(* IEC 61131-3 sources: daoli-st-library/DL_Algo (part 23) *)

(* ---- FB_DL_TriangleGenerator.st ---- *)
(*
  FB_DL_TriangleGenerator  —  三角波发生（相位连续 + 幅值/频率引脚化）/ Triangle wave generator
  分类 Category : DL_Algo
  码位 Code     : 16#02_3_87
  段位说明      : 86 格由 FB_DL_FrequencyGenerator 启用，本件启用相邻 87 格（一件一码）
  版本 Version  : 1.0.0
  来源 Source   : t2-1-lgf-siggen — 信号发生族第三基本波形（Sine/Sawtooth 同族）
  溯源 Origin   : clean-room 实现，相位累加三角波为公开经典方法，未复制任何源码行
  功能 Function : 1) 三角波发生：相位累加器在 [0,1) 内推进，方向标志交替升/降，
                  归一化输出 fNorm ∈ [0,1]，工程输出 fOut = fOffset + fAmplitude * (2*fNorm − 1)；
                  2) bPhaseReset 上升沿强制相位归零且方向置升（多路同相启动）；
                  3) fFreqHz = 0 时冻结在当前相位值（静止保持，不清输出）；
                  4) 波形形状按矩阵组纪律独立成件，明文禁用 eWaveform 枚举合并
                  （与 FB_DL_SineGenerator / 锯齿族分工，本件只做三角）。
  边界 Boundary : ① 幅值允许负值（输出相位反转语义：负幅值 = 倒相），非有限防御保持上次有效值；
                  ② 偏移 fOffset 非有限防御保持上次有效值；首扫按默认值；
                  ③ 无 TON/边沿实例：相位累加器法，任务周期由调用方经 tSampleTime 注入，
                  < T#10MS 钳位（与 FB_DL_RateLimiter 同口径）；
                  ④ 频率上限钳位（奈奎斯特防御）：高于任务频率一半时波形失真，越限按上限执行并置信息码；
                  ⑤ 方向切换在同一拍完成：fPhase >= 1 时先翻转方向再截去进位，避免相位突变尖峰。
  依赖 Depends  : 仅 Standard.library；与 FB_DL_SineGenerator（已注册）仅引脚口径对齐，不实例化
  码表 Error codes（本件格 02_3_87，子码步进 +0x100）:
    16#0002_0187 信息级：频率越上限已钳位（奈奎斯特防御，输出按钳后频率执行）
    16#0002_0287 信息级：相位复位沿生效（fPhase 归零、方向置升）
    16#0002_0387 信息级：非有限参数防御触发（保持上次有效值继续运行）

  修订历史 Revision :
    2026-11-19  v1.0.0  R39 首版（批次 1 · 序号 5）
*)

FUNCTION_BLOCK FB_DL_TriangleGenerator
VAR_INPUT
    bEnable     : BOOL := FALSE;      // 使能，FALSE 时冻结相位与输出 [-] / Enable, FALSE freezes phase and output
    fFreqHz     : REAL := 1.0;        // 目标频率 [Hz]，域 (0, 上限]，越限钳位 / Target frequency [Hz], clamped
    fAmplitude  : REAL := 100.0;      // 幅值 [EU]，可负（倒相语义），非有限保持 / Amplitude [EU], negative inverts phase
    fOffset     : REAL := 0.0;        // 直流偏移 [EU]，非有限保持 / DC offset [EU]
    bPhaseReset : BOOL := FALSE;      // 相位复位，上升沿相位归零、方向置升 / Phase reset, rising edge zeroes phase
    tSampleTime : TIME := T#100MS;    // 任务周期注入 [ms]，< T#10MS 钳位 / Task cycle time injected by caller
END_VAR
VAR_OUTPUT
    fOut        : REAL;               // 三角波工程输出 [EU] / Triangle engineering output [EU]
    fNormOut    : REAL;               // 归一化输出 [无量纲 0..1]，0 = 谷 / Normalized output, 0 = valley
    bRising     : BOOL;               // 本拍处于上升半周 [-] / Currently in the rising half-cycle
    uCycleCnt   : UDINT;              // 完整周期计数 [次]，降→升切换计一次，饱和 / Full cycle count, saturating
    bError      : BOOL;               // 故障标志，本件全信息级恒 FALSE（R21：信息级码不置故障）[-] / Fault flag, always FALSE, all codes info level
    uErrorId    : UDINT;              // 事件码，0 = 无事件（本件码均瞬时逐拍重算）/ Event code, transient, recomputed each scan
END_VAR
VAR
    rtPhaseReset : R_TRIG;            // 相位复位沿实例，主体首部无条件刷新 / Phase reset edge instance
    _fPhase      : REAL := 0.0;       // 内部相位累加器 [无量纲 0..1) / Internal phase accumulator
    _bUp         : BOOL := TRUE;      // 内部方向标志，TRUE = 升半周 / Internal direction flag, TRUE = rising
    _fFreqEff    : REAL := 1.0;       // 钳位后的生效频率 [Hz] / Clamped effective frequency
    _fAmpEff     : REAL := 100.0;     // 生效幅值 [EU] / Effective amplitude
    _fOffEff     : REAL := 0.0;       // 生效偏移 [EU] / Effective offset
    _fDt         : REAL := 0.1;       // 生效任务周期 [s] / Effective cycle time in seconds
    _fFreqLast   : REAL := 1.0;       // 上次有效频率保持载体 [Hz] / Last valid frequency hold carrier
    _fAmpLast    : REAL := 100.0;     // 上次有效幅值保持载体 [EU] / Last valid amplitude hold carrier
    _fOffLast    : REAL := 0.0;       // 上次有效偏移保持载体 [EU] / Last valid offset hold carrier
    _fNorm       : REAL := 0.0;       // 归一化中间量 [无量纲 0..1] / Normalized working value
    _bDefend     : BOOL;              // 本拍非有限防御触发标志 / Non-finite defense triggered this cycle
END_VAR
VAR CONSTANT
    DL_TG_DT_MIN     : TIME := T#10MS;      // 任务周期下限钳位 [ms] / Cycle time lower clamp
    DL_TG_FREQ_MAX   : REAL := 5.0;         // 频率组态上限（奈奎斯特防御，按 100ms 任务口径）[Hz] / Frequency configuration bound
    DL_TG_INF_CAP    : REAL := 1.0E30;      // 非有限值筛查幅值上限 / Non-finite magnitude screening cap
    DL_TG_CNT_MAX    : UDINT := 16#FFFF_FFFE;  // 周期计数饱和上限 [次] / Cycle count saturation bound
END_VAR

(* —— 段 0：边沿实例无条件周期刷新（R7 红线：严禁置于 IF/CASE 分支内） —— *)
rtPhaseReset(CLK := bPhaseReset);       // 相位复位沿刷新，每拍必调

(* —— 段 1：单拍量预清零 —— *)
uErrorId := 16#0000_0000;               // 事件码每拍重算（本件全信息级）
_bDefend := FALSE;                      // 防御标志预清零

(* —— 段 2：非有限防御与参数钳位（NaN/Inf 保持上次有效值） —— *)
IF (fFreqHz <> fFreqHz) OR (ABS(fFreqHz) > DL_TG_INF_CAP) OR ((fFreqHz - fFreqHz) <> 0.0) THEN
    _fFreqEff := _fFreqLast;            // 频率非有限：保持上次有效
    _bDefend := TRUE;
ELSE
    _fFreqLast := fFreqHz;
    IF fFreqHz < 0.0 THEN
        _fFreqEff := 0.0;               // 负频率钳零（冻结在当前相位值）
    ELSIF fFreqHz > DL_TG_FREQ_MAX THEN
        _fFreqEff := DL_TG_FREQ_MAX;    // 越上限钳位（奈奎斯特防御）
        uErrorId := 16#0002_0187;       // 信息级：频率已钳位
    ELSE
        _fFreqEff := fFreqHz;           // 域内直通
    END_IF
END_IF
IF (fAmplitude <> fAmplitude) OR (ABS(fAmplitude) > DL_TG_INF_CAP) OR ((fAmplitude - fAmplitude) <> 0.0) THEN
    _fAmpEff := _fAmpLast;              // 幅值非有限：保持上次有效
    _bDefend := TRUE;
ELSE
    _fAmpLast := fAmplitude;
    _fAmpEff := fAmplitude;             // 幅值允许负值（倒相语义），不钳位
END_IF
IF (fOffset <> fOffset) OR (ABS(fOffset) > DL_TG_INF_CAP) OR ((fOffset - fOffset) <> 0.0) THEN
    _fOffEff := _fOffLast;              // 偏移非有限：保持上次有效
    _bDefend := TRUE;
ELSE
    _fOffLast := fOffset;
    _fOffEff := fOffset;                // 偏移直通
END_IF
IF _bDefend THEN
    uErrorId := 16#0002_0387;           // 信息级：非有限防御触发（覆盖钳位码，防御码优先）
END_IF

(* —— 段 3：任务周期换算（与 FB_DL_RateLimiter 同口径：< T#10MS 钳位） —— *)
IF tSampleTime < DL_TG_DT_MIN THEN
    _fDt := 0.01;                       // 非法周期钳位 0.01 s
ELSE
    _fDt := TIME_TO_REAL(tSampleTime) / 1000.0;   // TIME 换算秒（显式标准转换）
END_IF

(* —— 段 4：相位复位沿（先于推进处理） —— *)
IF rtPhaseReset.Q THEN
    _fPhase := 0.0;                     // 相位归零
    _bUp := TRUE;                       // 方向置升
    uErrorId := 16#0002_0287;           // 信息级：相位复位生效（覆盖防御码，复位意图优先显式）
END_IF

(* —— 段 5：相位推进与方向翻转（失能冻结；频率 0 冻结在当前值） —— *)
IF bEnable AND (_fFreqEff > 0.0) THEN
    _fPhase := _fPhase + _fFreqEff * _fDt;      // 相位推进 = 频率 × 周期
    IF _fPhase >= 1.0 THEN
        _fPhase := _fPhase - 1.0;               // 截去进位（同拍完成，避免相位突变尖峰）
        IF _bUp THEN
            _bUp := FALSE;                      // 升满翻降（峰点换向）
        ELSE
            _bUp := TRUE;                       // 降满翻升（谷点换向）
            uCycleCnt := uCycleCnt + 1;         // 完整周期计数（降→升切换口径）
            IF uCycleCnt >= DL_TG_CNT_MAX THEN
                uCycleCnt := DL_TG_CNT_MAX;     // 计数饱和防回绕
            END_IF
        END_IF
        IF _fPhase >= 1.0 THEN
            _fPhase := 0.0;                     // 极端钳位兜底（频率越限多周回绕）
        END_IF
    END_IF
END_IF

(* —— 段 6：波形合成（升半周 fNorm = fPhase，降半周 fNorm = 1 − fPhase） —— *)
IF _bUp THEN
    _fNorm := _fPhase;                          // 上升半周：归一化随相位升
ELSE
    _fNorm := 1.0 - _fPhase;                    // 下降半周：归一化随相位降
END_IF
fNormOut := _fNorm;                             // 归一化镜像输出
fOut := _fOffEff + _fAmpEff * (2.0 * _fNorm - 1.0);   // 工程输出 = 偏移 + 幅值 ×（2·归一化 − 1）
bRising := _bUp AND bEnable;                    // 上升半周指示（失能时恒 FALSE）
bError := FALSE;                                // 本件全信息级：故障位恒 FALSE（R21）

END_FUNCTION_BLOCK

(* ---- FB_DL_TwoDofPid.st ---- *)
(*
  ==================================================================
  组件名 Component  : FB_DL_TwoDofPid
  分类   Category   : DL_Algo
  复杂度 Complexity  : cx4
  版本   Version    : 1.0.1
  功能   Purpose    : 二自由度 PID（设定值加权 beta / gamma），位置式：
                      u = Kp·(beta·sp - pv) + I + Kp·Td·(gamma·dsp/dt - dpv/dt)（滤后）。
                      积分作用于全误差 (sp - pv)；微分先行经 nFilter 一阶低通；
                      抗积分饱和（输出限幅方向与误差同向时停积分）；手动/自动
                      无扰切换（手动相把积分项跟踪为 fManOut - P - D）。
  来源   Source     : t2-5-modpid（参数域 beta / gamma）
  溯源   Origin     : IEC 61131-3 标准语义的道莅防御性实现；二自由度 PID 结构为
                      公开控制理论结果（Araki 参考跟踪 / 扰动抑制双自由度组织），
                      clean-room 自研实现，未复制任何闭源代码行。
  平台   Platform   : 纯 IEC 61131-3（LREAL 运算，无私有库、无幂运算符）
  作者   Author     : 道莅代码库 · PLC 编程专家（R56）
  ------------------------------------------------------------------
  边界 Boundary     :
                      一 本件只算控制器输出，不驱动执行器、不做自整定（属主边界）；
                      二 同拍双窗说明（R100）：本件无同拍双 TON 结构，微分滤波为一阶
                         差分实现，无定时器实例；
                      三 fTi <= 0 时积分项关闭（纯 PD 口径），fTd <= 0 时微分项关闭；
                      四 bInvalid = TRUE 时输出冻结保持末值（R191 显式声明，降级不静默）；
                      五 故障锁存（组态非法）解除路径 = bReset 上升沿（唯一路径，R188）；
                      六 无全局变量、无外部变量声明、无物理地址寻址、无定时器实例。
  输出契约 Output contract:
                      fOut 恒被钳在 [fOutMin, fOutMax]；bSatHi / bSatLo 为本拍限幅指示；
                      eFault 为锁存回放（eCfgIllegal 组态非法 / eInputBad 本拍输入非有限）。
  修订记录 Revision  :
    2026-11-20  v1.0.0  R56 首版（批 2 · 序号 8）
    2026-11-21  v1.0.1  R57 返修：手动相入口补 fManOut 有限性闸，无效拍冻结早退不进跟踪式
  ==================================================================
*)

TYPE E_DL_TdpFault :
(
    eNone     := 0, // 无成因 / no cause
    eCfgIllegal := 1, // 组态非法：增益或限幅越域（故障级，与 bError 配对）/ illegal config, gain or limit out of domain
    eInputBad := 2  // 本拍设定值或过程量非有限（信息级，输出冻结保持）/ the setpoint or process value is non finite this scan, the output holds frozen
);
END_TYPE

FUNCTION_BLOCK FB_DL_TwoDofPid
VAR_INPUT
    bAuto    : BOOL := TRUE;     // 自动模式，假 = 手动（无扰切换）[-] / auto mode, false is manual with a bumpless transfer
    bReset   : BOOL := FALSE;    // 复位上升沿清故障锁存与积分 [-] / reset rising edge clears the fault latch and the integral
    fSp      : LREAL := 0.0;     // 设定值 [工程单位] / setpoint [engineering unit]
    fPv      : LREAL := 0.0;     // 过程量实测 [工程单位] / measured process value [engineering unit]
    fManOut  : LREAL := 0.0;     // 手动输出值 [工程单位] / manual output value [engineering unit]
    fKp      : LREAL := 1.0;     // 比例增益，域 大于零 / proportional gain, domain above zero
    fTi      : LREAL := 10.0;    // 积分时间 [秒]，0 = 积分关闭 / integral time [second], zero disables the integral
    fTd      : LREAL := 0.0;     // 微分时间 [秒]，0 = 微分关闭 / derivative time [second], zero disables the derivative
    fBeta    : LREAL := 1.0;     // 设定值比例加权（抑超调自由度），域 0..1 / setpoint proportional weight [dimensionless], domain zero to one
    fGamma   : LREAL := 0.0;     // 设定值微分加权，域 0..1 / setpoint derivative weight, domain zero to one
    nFilter  : INT := 10;        // 微分低通系数 n（Td/n 为滤波时间），域 1..100 / derivative low pass coefficient n, domain one to one hundred
    fOutMin  : LREAL := 0.0;     // 输出下限 [工程单位] / output floor [engineering unit]
    fOutMax  : LREAL := 100.0;   // 输出上限 [工程单位]，域 大于下限 / output ceiling [engineering unit], above the floor
    fDtS     : LREAL := 0.01;    // 调用周期 [秒]，域 大于零 / call period [second], domain above zero
END_VAR
VAR_OUTPUT
    fOut     : LREAL := 0.0;   // 控制器输出 [工程单位] / controller output [engineering unit]
    bSatHi   : BOOL := FALSE;  // 本拍输出顶上限 [-] / the output hit the ceiling this scan
    bSatLo   : BOOL := FALSE;  // 本拍触下限 [-] / the output hit the floor this scan
    bInvalid : BOOL := FALSE;  // 本拍输出无效（冻结保持末值）[-] / the outlet is void this scan, the last value holds frozen
    eFault   : E_DL_TdpFault := E_DL_TdpFault.eNone; // 成因出口，锁存回放 [枚举] / cause outlet replayed from the latch [enum]
    bError   : BOOL := FALSE;  // 故障锁存标志 [-] / fault latch flag
END_VAR
VAR
    rtReset  : R_TRIG;  // 复位沿检测，段 0 无条件刷新 / reset edge, refreshed unconditionally in segment zero
    _eFaulC  : E_DL_TdpFault := E_DL_TdpFault.eNone; // 故障级成因，锁存至复位沿 / fault cause, latched until the reset edge
    _bFault  : BOOL := FALSE; // 故障锁存位 [-] / fault latch bit
    _bInit   : BOOL := FALSE; // 首扫初始化完成标志（R310）/ first scan initialisation flag
    _bInOk   : BOOL := FALSE; // 本拍 sp / pv 均有限 [-] / both sp and pv are finite this scan
    _fI      : LREAL := 0.0;  // 积分项保持量 [工程单位] / the integral term holder [engineering unit]
    _fDfilt  : LREAL := 0.0;  // 微分滤波保持量 [工程单位] / the derivative filter holder [engineering unit]
    _fPvPrev : LREAL := 0.0;  // 上拍过程量快照 [工程单位] / previous scan process value snapshot [engineering unit]
    _fSpPrev : LREAL := 0.0;  // 上拍设定值快照 [工程单位] / previous scan setpoint snapshot [engineering unit]
    _fP      : LREAL := 0.0;  // 本拍比例项 [工程单位] / the proportional term this scan [engineering unit]
    _fDraw   : LREAL := 0.0;  // 微分原始量 [工程单位] / the raw derivative term [engineering unit]
    _fE      : LREAL := 0.0;  // 全误差（sp - pv）[工程单位] / the full error [engineering unit]
    _fUPre   : LREAL := 0.0;  // 限幅前输出 [工程单位] / the pre clamp output [engineering unit]
    _fFiltB  : LREAL := 0.0;  // 微分滤波权（dt/(dt+Td/n)）[无量纲] / the derivative filter weight
END_VAR

// 段 0｜沿检测无条件周期刷新（禁入分支）/ segment 0, unconditional refresh of the edge detector
rtReset(CLK := bReset); // 复位沿无条件刷新 / unconditional refresh of the reset edge

// 段 1｜首扫初始化（R310）：快照与积分从确定起点起步 / segment 1, first scan initialisation
IF NOT _bInit THEN // 首扫一拍 / the very first scan
    _bInit := TRUE; // 置首扫完成标志 / raise the first scan flag
    _eFaulC := E_DL_TdpFault.eNone; // 故障级成因清零 / clear the fault cause
    _bFault := FALSE; // 故障锁存清零 / clear the fault latch
    _fI := 0.0; // 积分项清零 / clear the integral term
    _fDfilt := 0.0; // 微分滤波清零 / clear the derivative filter
    _fPvPrev := fPv; // 快照取当拍 / the snapshot takes this scan
    _fSpPrev := fSp; // 快照取当拍 / the snapshot takes this scan
END_IF

// 段 2｜复位沿作用域：清锁存 / 清积分与滤波（快照同步归位，三项逐项声明）/ segment 2, reset edge scope declared item by item
IF rtReset.Q THEN // 复位沿 / the reset edge
    _bFault := FALSE; // 作用域一：清故障锁存 / scope one, clear the fault latch
    _eFaulC := E_DL_TdpFault.eNone; // 作用域一：清故障级成因 / scope one, clear the fault cause
    _fI := 0.0; // 作用域二：清积分项 / scope two, clear the integral term
    _fDfilt := 0.0; // 作用域二：清微分滤波 / scope two, clear the derivative filter
    _fPvPrev := fPv; // 作用域三：快照归位 / scope three, the snapshot parks
    _fSpPrev := fSp; // 作用域三：快照归位 / scope three, the snapshot parks
END_IF

// 段 3｜组态域闸（R151 全覆盖）/ segment 3, configuration domain gate over every parameter pin
IF (fKp <= 0.0) OR (fKp <> fKp) OR ((fKp - fKp) <> (fKp - fKp)) OR (fTi < 0.0) OR (fTi <> fTi) OR (fTd < 0.0) OR (fTd <> fTd) OR (fBeta < 0.0) OR (fBeta > 1.0) OR (fBeta <> fBeta) OR (fGamma < 0.0) OR (fGamma > 1.0) OR (fGamma <> fGamma) OR (nFilter < 1) OR (nFilter > 100) OR (fOutMax <= fOutMin) OR (fOutMax <> fOutMax) OR (fDtS <= 0.0) OR (fDtS <> fDtS) THEN // 任一参数越域或非有限 / any parameter out of domain or non finite
    IF (NOT _bFault) AND (_eFaulC = E_DL_TdpFault.eNone) THEN // 未锁存才迁移（防同拍抹除）/ migrate only while unlatched
        _bFault := TRUE; // 置故障锁存 / raise the fault latch
        _eFaulC := E_DL_TdpFault.eCfgIllegal; // 故障级成因（R45 配对 bError）/ the fault cause paired with bError
    END_IF
END_IF

// 段 4｜输入有限性闸与冻结语义 / segment 4, the input finiteness gate and the frozen semantics
_bInOk := (fSp = fSp) AND ((fSp - fSp) = (fSp - fSp)) AND (fPv = fPv) AND ((fPv - fPv) = (fPv - fPv)); // sp / pv 有限性 / finiteness of sp and pv

// 段 5｜无扰切换：手动相把积分项跟踪为 fManOut - P - D / segment 5, the bumpless transfer, the manual phase tracks the integral
IF NOT bAuto THEN // 手动相 / the manual phase
    IF (fManOut <> fManOut) OR ((fManOut - fManOut) <> (fManOut - fManOut)) THEN // 手动输出非有限（x<>x 判 NaN，x-x<>x-x 判 Inf，v1.0.1 返修）/ the manual output is non finite (v1.0.1 fix)
        IF NOT _bFault THEN // 故障锁存优先回放，信息级不覆盖故障码 / the fault latch replays first, an informational cause never overwrites a fault code
            _eFaulC := E_DL_TdpFault.eInputBad; // 信息级成因（R45 不配对 bError）/ the informational cause, not paired with bError
        END_IF
        bInvalid := TRUE; // 置无效标志 / raise the invalid flag
        bSatHi := FALSE; // 限幅指示为假 / the saturation flags are false
        bSatLo := FALSE; // 限幅指示为假 / the saturation flags are false
        eFault := _eFaulC; // 成因出口锁存回放 / the cause outlet replayed from the latch
        bError := _bFault; // 故障标志与锁存位同源 / the fault flag shares the latch source
        _fPvPrev := fPv; // 快照推进（防恢复时微分踢）/ advance the snapshot against a derivative kick
        _fSpPrev := fSp; // 快照推进 / advance the snapshot
        RETURN; // 早退，fOut 冻结保持末值，不进跟踪式（R191 已声明）/ early return, fOut holds frozen, no tracking (R191 declared)
    END_IF
    _fP := fKp * (fBeta * fSp - fPv); // 比例项同口径计算（为跟踪做准备）/ the proportional term for the tracking base
    _fI := fManOut - _fP - _fDfilt; // 积分项跟踪，自动恢复时无扰 / the integral tracks for a bumpless auto resume
    fOut := fManOut; // 手动输出直通 / the manual output passes through
    IF fOut > fOutMax THEN // 手动输出上钳 / clamp the manual output high
        fOut := fOutMax; // 钳到上限 / clamp to the ceiling
    ELSIF fOut < fOutMin THEN // 手动输出下钳 / clamp the manual output low
        fOut := fOutMin; // 钳到下限 / clamp to the floor
    END_IF
    bSatHi := FALSE; // 手动相限幅指示为假 / the saturation flags are false in manual
    bSatLo := FALSE; // 手动相限幅指示为假 / the saturation flags are false in manual
    bInvalid := (NOT _bInOk) OR _bFault; // 有效性随输入与锁存 / the validity follows the input and the latch
    eFault := _eFaulC; // 成因出口锁存回放 / the cause outlet replayed from the latch
    bError := _bFault; // 故障标志与锁存位同源 / the fault flag shares the latch source
    _fPvPrev := fPv; // 快照推进 / advance the snapshot
    _fSpPrev := fSp; // 快照推进 / advance the snapshot
    RETURN; // 手动相早退（出口段已完整施加，R94）/ the manual phase early return with a complete outlet
END_IF

// 段 6｜自动相：无效输入冻结保持 / segment 6, the auto phase, a void input holds frozen
IF (NOT _bInOk) OR _bFault THEN // 输入无效或故障锁存 / the input is void or faulted
    IF (NOT _bInOk) AND (NOT _bFault) THEN // 输入缺陷才记信息级成因（不覆盖故障码）/ only an input defect records the informational cause, never over a fault latch
        _eFaulC := E_DL_TdpFault.eInputBad; // 信息级成因，每拍重算 / the informational cause, recomputed every scan
    END_IF
    bInvalid := TRUE; // 置无效标志 / raise the invalid flag
    bSatHi := FALSE; // 限幅指示为假 / the saturation flags are false
    bSatLo := FALSE; // 限幅指示为假 / the saturation flags are false
    eFault := _eFaulC; // 成因出口锁存回放 / the cause outlet replayed from the latch
    bError := _bFault; // 故障标志与锁存位同源 / the fault flag shares the latch source
    _fPvPrev := fPv; // 快照推进（防恢复时微分踢）/ advance the snapshot against a derivative kick
    _fSpPrev := fSp; // 快照推进 / advance the snapshot
    RETURN; // 早退，fOut 冻结保持末值（R191 已在头注释声明）/ early return, fOut holds frozen per the declared semantics
END_IF

// 段 7｜比例与微分先行（幂次无，显式乘法）/ segment 7, the proportional and the derivative lead terms
_fE := fSp - fPv; // 全误差 / the full error
_fP := fKp * (fBeta * fSp - fPv); // 加权比例项 / the weighted proportional term
IF fTd > 0.0 THEN // 微分开启 / the derivative is on
    _fDraw := fTd * (fGamma * (fSp - _fSpPrev) - (fPv - _fPvPrev)) / fDtS; // 加权微分原始量，除子为周期已证大于零 / the weighted raw derivative, the divisor is the proven period
    _fFiltB := fDtS / (fDtS + fTd / INT_TO_LREAL(nFilter)); // 一阶低通权，除子已证大于零 / the first order weight with a proven divisor
    _fDfilt := _fDfilt + _fFiltB * (_fDraw - _fDfilt); // 微分低通推进 / advance the derivative low pass
ELSE // 微分关闭 / the derivative is off
    _fDfilt := 0.0; // 微分项归零 / the derivative term is zeroed
END_IF

// 段 8｜积分与抗饱和：先算限幅前输出，再按方向条件积分 / segment 8, the integral with anti windup, the clamp direction gates the accumulation
_fUPre := _fP + _fI + _fDfilt; // 限幅前输出 / the pre clamp output
IF (fTi > 0.0) THEN // 积分开启 / the integral is on
    IF NOT ((_fUPre > fOutMax) AND (_fE > 0.0)) AND NOT ((_fUPre < fOutMin) AND (_fE < 0.0)) THEN // 输出未沿误差方向饱和才积分（抗 windup）/ the integration only runs when the output is not saturated in the error direction
        _fI := _fI + (fKp / fTi) * _fE * fDtS; // 积分推进，除子为积分时间已证大于零 / the integral step with the proven divisor
    END_IF
END_IF
_fUPre := _fP + _fI + _fDfilt; // 积分后重算限幅前输出 / recompute after the integral

// 段 9｜限幅与限幅指示 / segment 9, the clamp and the saturation flags
bSatHi := FALSE; // 限幅指示预置假 / preset the saturation flags to false
bSatLo := FALSE; // 限幅指示预置假 / preset the saturation flags to false
IF _fUPre > fOutMax THEN // 顶上限 / above the ceiling
    fOut := fOutMax; // 钳到上限 / clamp to the ceiling
    bSatHi := TRUE; // 置顶上限指示 / raise the ceiling flag
ELSIF _fUPre < fOutMin THEN // 触下限 / below the floor
    fOut := fOutMin; // 钳到下限 / clamp to the floor
    bSatLo := TRUE; // 置触下限指示 / raise the floor flag
ELSE // 域内 / inside the domain
    fOut := _fUPre; // 直接出口 / straight to the outlet
END_IF

// 段 10｜快照推进与统一出口 / segment 10, the snapshot advance and the unified outlet
_fPvPrev := fPv; // 过程量快照推进 / advance the process snapshot
_fSpPrev := fSp; // 设定值快照推进 / advance the setpoint snapshot
IF (_eFaulC = E_DL_TdpFault.eInputBad) AND (NOT _bFault) THEN // 输入已恢复 / the input has recovered
    _eFaulC := E_DL_TdpFault.eNone; // 信息级成因随恢复撤销 / the informational cause is revoked on recovery
END_IF
bInvalid := FALSE; // 自动有效拍 / the valid auto scan
eFault := _eFaulC; // 成因出口锁存回放 / the cause outlet replayed from the latch
bError := _bFault; // 故障标志与锁存位同源 / the fault flag shares the latch source
END_FUNCTION_BLOCK

(* ---- FB_DL_UvDoseCtrl.st ---- *)
(*
  ==================================================================
  组件名 Component  : FB_DL_UvDoseCtrl
  分类   Category   : DL_Algo
  复杂度 Complexity  : cx5
  版本   Version    : 1.0.0
  功能   Purpose    : UV 剂量控制。剂量 = 光强 × 曝晒时间（D = ∫I·kLamp·dt），
                      按剩余剂量误差 PI 闭环调光强输出（0..100%），累计达目标置
                      bDoseDone 单拍脉冲；灯管老化补偿系数 kLamp 外部给定；光强
                      非有限 / 负值闸；累计溢出保护；满输出长期照度不足判
                      eLampWeak；过冲超容差判 eDoseOvershoot。
  来源   Source     : 自研线（公开物理定义：剂量 = 强度 × 时间积分）
  溯源   Origin     : IEC 61131-3 标准语义的道莅防御性实现；UV 剂量定义为公开
                      光化学语义，clean-room 自研实现，未复制任何闭源代码行。
  平台   Platform   : 纯 IEC 61131-3（TON / R_TRIG / LREAL，无私有库）
  作者   Author     : 道莅代码库 · PLC 编程专家（R56）
  ------------------------------------------------------------------
  边界 Boundary     :
                      一 本件只算调光输出与剂量累计，不驱动灯管电源本体（属主边界）；
                      二 bRun = FALSE 时调光输出归零、累计冻结保持（R191 显式声明）；
                      三 剂量累计溢出保护：累计达 1.0E9 mJ/cm² 上限即饱和（远超
                         任何工艺目标，防长跑溢出，R63 反算：1.0E9 在 LREAL 精确可表）；
                      四 故障锁存解除路径 = bReset 上升沿（唯一路径，R188）；
                      五 无全局变量、无外部变量声明、无物理地址寻址。
  输出契约 Output contract:
                      fDimPct 恒在 [0, 100]；fDoseAcc 为累计剂量 [毫焦每平方厘米]；
                      bDoseDone 为单拍脉冲（内部 _bDoneInt 置位、统一出口映射后撤销，
                      R187 两段式）；eFault 为锁存回放；
                      ePhaseBad 为非法相位兜底专用成员（R128）。
  修订记录 Revision  :
    2026-11-20  v1.0.0  R56 首版（批 4 · 序号 17）
  ==================================================================
*)

TYPE E_DL_UdcPhase :
(
    eIdle  := 0,  // 空闲：等运行电平 / idle, waiting for the run level
    eDose  := 10, // 照射：闭环调光与剂量累计 / dosing, the closed loop dimming and the accumulation
    eDone  := 20, // 达标：脉冲已出，灯关驻留 / done, the pulse was raised and the lamp is off
    eFault := 90  // 故障：成因锁存，灯关 / fault, the cause is latched with the lamp off
);
END_TYPE

TYPE E_DL_UdcFault :
(
    eNone          := 0, // 无成因 / no cause
    eLampWeak      := 1, // 满输出照度不足（灯管老化，故障级，与 bError 配对）/ the intensity is weak at a full output, an aged lamp, fault grade paired with bError
    eDoseOvershoot := 2, // 剂量过冲超容差（故障级，与 bError 配对）/ the dose overshot the tolerance, fault grade paired with bError
    eSensorBad     := 3, // 光强非有限或负值（故障级，与 bError 配对）/ the intensity is non finite or negative, fault grade paired with bError
    ePhaseBad      := 4  // 非法相位兜底（故障级，与 bError 配对）/ illegal phase fallback, fault grade paired with bError
);
END_TYPE

FUNCTION_BLOCK FB_DL_UvDoseCtrl
VAR_INPUT
    bEnable    : BOOL := TRUE;    // 使能，失能时停判级回空闲 [-] / enable, the grading stops when disabled
    bReset     : BOOL := FALSE;   // 复位上升沿清故障锁存并剂量归零重批 [-] / reset rising edge clears the latch and zeroes the dose for a fresh batch
    bRun       : BOOL := FALSE;   // 运行电平，真 = 曝晒窗开 [-] / the run level, true opens the exposure window
    fIntensity : LREAL := 0.0;    // 光强实测 [毫瓦每平方厘米] / the measured intensity [milliwatt per square centimetre]
    fDoseTarget: LREAL := 100.0;  // 目标剂量 [毫焦每平方厘米]，域 大于零 / the target dose [millijoule per square centimetre], domain above zero
    kLamp      : LREAL := 1.0;    // 灯管老化补偿系数（有效光强占比），域 0..1 / the lamp ageing compensation factor, domain zero to one
    fKp        : LREAL := 5.0;    // PI 比例增益 [百分比每毫焦] / the PI proportional gain [percent per millijoule]
    fKi        : LREAL := 0.5;    // PI 积分增益 [百分比每毫焦每秒] / the PI integral gain
    fIntMin    : LREAL := 5.0;    // 最小有效照度 [毫瓦每平方厘米]，域 大于零 / the minimum effective intensity, domain above zero
    fOverTolPct: LREAL := 5.0;    // 过冲容差 [百分比]，域 大于零 / the overshoot tolerance [percent], domain above zero
    tWeakTo    : TIME := T#30S;   // 灯弱确认窗 [毫秒]，域 大于零 / the weak lamp confirm window [millisecond], domain above zero
    fDtS       : LREAL := 0.1;    // 调用周期 [秒]，域 大于零 / the call period [second], domain above zero
END_VAR
VAR_OUTPUT
    fDimPct   : LREAL := 0.0;  // 调光输出 [百分比] / the dimming output [percent]
    bDoseDone : BOOL := FALSE; // 剂量达标单拍脉冲 [-] / the dose done single shot pulse
    fDoseAcc  : LREAL := 0.0;  // 累计剂量 [毫焦每平方厘米] / the accumulated dose [millijoule per square centimetre]
    ePhase    : E_DL_UdcPhase := E_DL_UdcPhase.eIdle; // 相位出口 [枚举] / phase outlet [enum]
    eFault    : E_DL_UdcFault := E_DL_UdcFault.eNone; // 成因出口，锁存回放 [枚举] / cause outlet replayed from the latch [enum]
    bError    : BOOL := FALSE; // 故障锁存标志 [-] / fault latch flag
END_VAR
VAR
    rtReset  : R_TRIG; // 复位沿检测，段 0 无条件刷新 / reset edge, refreshed unconditionally in segment zero
    tonWeak  : TON;    // 灯弱确认窗，段 0 无条件刷新 / the weak lamp window, refreshed unconditionally
    _ePhase  : E_DL_UdcPhase := E_DL_UdcPhase.eIdle; // 内部相位，CASE 唯一写入目标 / internal phase, the only CASE write target
    _eFaulC  : E_DL_UdcFault := E_DL_UdcFault.eNone; // 故障级成因，锁存至复位沿 / fault cause, latched until the reset edge
    _bFault  : BOOL := FALSE; // 故障锁存位 [-] / fault latch bit
    _bInit   : BOOL := FALSE; // 首扫初始化完成标志（R310）/ first scan initialisation flag
    _bDoneInt: BOOL := FALSE; // 达标脉冲内部位，统一出口映射 / internal done bit, mapped at the unified outlet
    _bInOk   : BOOL := FALSE; // 光强有限且非负 [-] / the intensity is finite and non negative
    _bCfgOk  : BOOL := FALSE; // 组态参数域内 [-] / the configuration is inside the domain
    _bWeakRaw: BOOL := FALSE; // 满输出照度不足原始判据 [-] / the raw weak lamp verdict
    _fRate   : LREAL := 0.0;  // 剂量率 [毫焦每平方厘米每秒] / the dose rate
    _fE      : LREAL := 0.0;  // 剩余剂量误差 [毫焦每平方厘米] / the remaining dose error
    _fUPre   : LREAL := 0.0;  // 限幅前调光输出 [百分比] / the pre clamp dimming output
    _fI      : LREAL := 0.0;  // 积分项保持量 [百分比] / the integral term holder [percent]
    _fTol    : LREAL := 0.0;  // 过冲绝对容差 [毫焦每平方厘米] / the absolute overshoot tolerance
END_VAR

// 段 0｜定时器与沿检测无条件周期刷新（禁入分支），IN 只串相位闸与状态闸 / segment 0, unconditional refresh with the phase and state gates
rtReset(CLK := bReset); // 复位沿无条件刷新 / unconditional refresh of the reset edge
tonWeak(IN := _bWeakRaw AND (_ePhase = E_DL_UdcPhase.eDose) AND (NOT _bFault), PT := tWeakTo); // 灯弱确认窗，IN 串原始判据与相位闸 / the weak lamp window with the raw verdict and the phase gate

// 段 1｜首扫初始化（R310）/ segment 1, first scan initialisation
IF NOT _bInit THEN // 首扫一拍 / the very first scan
    _bInit := TRUE; // 置首扫完成标志 / raise the first scan flag
    _ePhase := E_DL_UdcPhase.eIdle; // 相位从空闲起步 / the phase starts from idle
    _eFaulC := E_DL_UdcFault.eNone; // 故障级成因清零 / clear the fault cause
    _bFault := FALSE; // 故障锁存清零 / clear the fault latch
    _fI := 0.0; // 积分项清零 / clear the integral term
    fDoseAcc := 0.0; // 剂量清零 / clear the dose
END_IF

// 段 2｜复位沿作用域：清锁存 / 迁相位 / 清剂量与积分（三项逐项声明）/ segment 2, reset edge scope declared item by item
IF rtReset.Q THEN // 复位沿 / the reset edge
    _bFault := FALSE; // 作用域一：清故障锁存 / scope one, clear the fault latch
    _eFaulC := E_DL_UdcFault.eNone; // 作用域一：清故障级成因 / scope one, clear the fault cause
    _ePhase := E_DL_UdcPhase.eIdle; // 作用域二：迁回空闲相 / scope two, migrate back to idle
    fDoseAcc := 0.0; // 作用域三：清剂量累计 / scope three, clear the dose accumulation
    _fI := 0.0; // 作用域三：清积分项 / scope three, clear the integral term
END_IF

// 段 3｜组态与输入域闸（R151 全覆盖）/ segment 3, the configuration and input domain gates
_bInOk := (fIntensity = fIntensity) AND ((fIntensity - fIntensity) = (fIntensity - fIntensity)) AND (fIntensity >= 0.0); // 光强有限且非负 / the intensity is finite and non negative
_bCfgOk := (fDoseTarget > 0.0) AND (fDoseTarget = fDoseTarget) AND (kLamp >= 0.0) AND (kLamp <= 1.0) AND (kLamp = kLamp) AND (fKp > 0.0) AND (fKp = fKp) AND (fKi >= 0.0) AND (fKi = fKi) AND (fIntMin > 0.0) AND (fIntMin = fIntMin) AND (fOverTolPct > 0.0) AND (fOverTolPct = fOverTolPct) AND (tWeakTo > T#0S) AND (fDtS > 0.0) AND (fDtS = fDtS); // 组态参数域判定 / the configuration domain verdict
IF (NOT _bInOk) OR (NOT _bCfgOk) THEN // 光强无效或组态非法 / a void intensity or an illegal configuration
    IF NOT _bFault THEN // 未锁存才迁移（防同拍抹除）/ migrate only while unlatched
        _bFault := TRUE; // 置故障锁存 / raise the fault latch
        _eFaulC := E_DL_UdcFault.eSensorBad; // 故障级成因（R45 配对 bError）/ the fault cause paired with bError
        _ePhase := E_DL_UdcPhase.eFault; // 迁故障相 / migrate to the fault phase
    END_IF
END_IF

// 段 4｜相位机：ENUM + CASE，含 ELSE 非法相位兜底（R128）/ segment 4, the phase machine with an ELSE fallback
CASE _ePhase OF
E_DL_UdcPhase.eIdle: // 空闲相：等运行电平 / the idle phase, waiting for the run level
    fDimPct := 0.0; // 灯关 / the lamp is off
    IF bEnable AND (NOT _bFault) AND bRun THEN // 运行电平受理 / the run level is accepted
        _fI := 0.0; // 积分项清零 / clear the integral term
        _ePhase := E_DL_UdcPhase.eDose; // 迁照射相 / migrate to the dose phase
    END_IF

E_DL_UdcPhase.eDose: // 照射相：闭环调光 + 剂量累计（退出条件 ≥2：达标 / 过冲 / 灯弱 / 失能 / 停运行，R98）/ the dose phase with at least two exit conditions
    IF NOT bEnable THEN // 失能 / disabled
        fDimPct := 0.0; // 灯关 / the lamp is off
        _ePhase := E_DL_UdcPhase.eIdle; // 回空闲相 / back to idle
    ELSIF NOT bRun THEN // 曝晒窗关：调光归零、累计冻结保持（R191 显式声明）/ the window closed, the dimming zeroes and the dose freezes
        fDimPct := 0.0; // 灯关 / the lamp is off
        _fI := 0.0; // 积分项清零（防恢复时积分踢）/ clear the integral against a kick on resume
    ELSE // 曝晒中 / exposing
        IF _bInOk AND _bCfgOk THEN // 输入与组态合法 / the input and the config are legal
            _fRate := fIntensity * kLamp; // 剂量率 = 光强 × 老化补偿系数 / the dose rate, the intensity times the factor
            fDoseAcc := fDoseAcc + _fRate * fDtS; // 剂量累计 / accumulate the dose
            IF fDoseAcc > 1.0E9 THEN // 累计溢出保护（饱和口径，R63 反算）/ the overflow protection with the saturation basis
                fDoseAcc := 1.0E9; // 饱和到上限 / saturate at the ceiling
            END_IF
            _fTol := fDoseTarget * fOverTolPct / 100.0; // 过冲绝对容差，除子为常量一百 / the absolute tolerance with the constant divisor
            _fE := fDoseTarget - fDoseAcc; // 剩余剂量误差 / the remaining dose error
            _fUPre := fKp * _fE + _fI; // 限幅前调光输出 / the pre clamp dimming output
            IF NOT ((_fUPre >= 100.0) AND (_fE > 0.0)) THEN // 未沿误差方向饱和才积分（抗 windup）/ the integration is gated against the saturation direction
                _fI := _fI + fKi * _fE * fDtS; // 积分推进 / the integral step
            END_IF
            _fUPre := fKp * _fE + _fI; // 积分后重算 / recompute after the integral
            IF _fUPre < 0.0 THEN // 下限钳零 / clamp the floor to zero
                fDimPct := 0.0; // 输出归零 / the output is zeroed
            ELSIF _fUPre > 100.0 THEN // 上限钳百 / clamp the ceiling to one hundred
                fDimPct := 100.0; // 输出满幅 / the output is full
            ELSE // 域内 / inside the domain
                fDimPct := _fUPre; // 直接出口 / straight to the outlet
            END_IF
            _bWeakRaw := (fDimPct >= 99.0) AND (_fRate < fIntMin); // 满输出照度不足原始判据 / the raw weak lamp verdict
            IF fDoseAcc > fDoseTarget + _fTol THEN // 过冲超容差（优先归因，R190 独立成因）/ the overshoot takes the cause priority
                _bFault := TRUE; // 置故障锁存 / raise the fault latch
                _eFaulC := E_DL_UdcFault.eDoseOvershoot; // 故障级成因（R45 配对 bError）/ the fault cause paired with bError
                _ePhase := E_DL_UdcPhase.eFault; // 迁故障相 / migrate to the fault phase
            ELSIF tonWeak.Q THEN // 灯弱确认窗到 / the weak lamp window elapsed
                _bFault := TRUE; // 置故障锁存 / raise the fault latch
                _eFaulC := E_DL_UdcFault.eLampWeak; // 故障级成因（R45 配对 bError）/ the fault cause paired with bError
                _ePhase := E_DL_UdcPhase.eFault; // 迁故障相 / migrate to the fault phase
            ELSIF fDoseAcc >= fDoseTarget THEN // 剂量达标 / the dose target is reached
                _bDoneInt := TRUE; // 达标脉冲内部位置位（统一出口映射，R187）/ raise the internal done bit
                _ePhase := E_DL_UdcPhase.eDone; // 迁达标相 / migrate to the done phase
            END_IF
        ELSE // 输入或组态非法：灯关防御 / a void input or config, the lamp is off as a defence
            fDimPct := 0.0; // 灯关 / the lamp is off
        END_IF
    END_IF

E_DL_UdcPhase.eDone: // 达标相：灯关驻留，等运行撤或复位 / the done phase, the lamp is off until the run drops or a reset
    fDimPct := 0.0; // 灯关 / the lamp is off
    IF (NOT bEnable) OR (NOT bRun) THEN // 失能或运行撤 / disabled or the run dropped
        _ePhase := E_DL_UdcPhase.eIdle; // 回空闲相 / back to idle
    END_IF

E_DL_UdcPhase.eFault: // 故障相：灯关，成因锁存，等复位沿 / the fault phase, the lamp is off until the reset edge
    fDimPct := 0.0; // 灯关（安全侧）/ the lamp is off, the safe side
    IF NOT bEnable THEN // 失能 / disabled
        _ePhase := E_DL_UdcPhase.eIdle; // 迁未使能相 / migrate to idle
    END_IF

ELSE // 非法相位兜底（R128）/ the illegal phase fallback
    _bFault := TRUE; // 置故障锁存 / raise the fault latch
    _eFaulC := E_DL_UdcFault.ePhaseBad; // 故障级成因（R45 配对 bError）/ the fault cause paired with bError
    _ePhase := E_DL_UdcPhase.eFault; // 迁故障相 / migrate to the fault phase
END_CASE

// 段 5｜统一出口 / segment 5, the unified outlet
bDoseDone := _bDoneInt; // 达标脉冲映射本拍值 / map the done pulse for this scan
_bDoneInt := FALSE; // 映射后立即撤销，保证单拍宽度（R187 两段式）/ revoke right after mapping
IF _bFault THEN // 故障锁存优先 / the fault latch takes priority
    eFault := _eFaulC; // 故障级成因锁存回放（R152）/ the fault cause replayed from the latch
ELSE
    eFault := E_DL_UdcFault.eNone; // 无锁存即无成因 / no latch, no cause
END_IF
ePhase := _ePhase; // 相位出口单点映射 / single point phase outlet mapping
bError := _bFault; // 故障标志与锁存位同源 / the fault flag shares the latch source
END_FUNCTION_BLOCK

(* ---- FB_DL_VavPressureReset.st ---- *)
(*
  FB_DL_VavPressureReset  —  VAV 静压重置（最不利末端阀位寻优 + 步长限幅） / VAV duct static-pressure reset by worst-case terminal damper optimisation with step limiting
  分类 Category : DL_Algo
  版本 Version  : 1.0.0
  来源 Source   : t1-2-oscat-building — 楼宇变风量静压重置算法族深化
  溯源 Origin   : 道莅 clean-room 实现；以最不利末端阀位为反馈的静压爬坡重置（死区 + 步长限幅）为公开 VAV 节能算法，未复制任何源码行
  功能 Function : 1) 偏差 _fErrPct = fDamperTargetPct - fWorstDamperPct（最不利末端阀位对目标阀位）；
                  2) 死区保持：|偏差| <= fDeadbandPct 时设定保持不变（不动作）；
                  3) 爬坡寻优：偏差为正（阀位偏小，需更大静压）每周期加 fStepKpa，
                  偏差为负每周期减 fStepKpa，单周期变化量恒等于步长（限速内置）；
                  4) 硬限幅：设定钳制到 [fSpMinKpa, fSpMaxKpa]，限幅后二次复核；
                  5) 本件只有故障码、无信息码（派单硬约束）。
  接口 Interface: 输入最不利阀位/目标阀位/死区/步长/上下限；输出静压设定与动作镜像
  边界 Boundary : ① 组态闸：fSpMaxKpa <= fSpMinKpa、fStepKpa <= 0.0、fDeadbandPct < 0.0、
                  fDamperTargetPct 不在 (0, 100) 开区间 → 0387 锁存；
                  ② 阀位与设定量非有限（NaN 自反 + Inf 差值自减）→ 0387 锁存，输出冻结保持
                  （本件为设定类算法，冻结保持不降级，语义已在头注释声明，R191）；
                  ③ 浮点判据全容差式，禁 = / <> 判等；④ 仅一个 R_TRIG 复位沿，段 0 无条件调用；
                  ⑤ 故障相迁出唯一路径 = bReset 上升沿；⑥ 零全局耦合（无 GVL / %I %Q %M）。
  依赖 Depends  : Standard.library（R_TRIG）
  码表 Error codes（Algo 段 0002，故障窗口 0387；本件无信息码）:
    16#0002_0387 故障级：VAV 静压重置故障总码（组态非法 / 阀位或设定非有限），
                 锁存至 bReset 上升沿；归因见 eCause，不新增码位（派单硬约束单码）
  修订历史 Revision :
    2026-11-19  v1.0.0  R43 首版（批次 3 · 序号 11）
*)

TYPE E_DL_VprState :
(
    eIdle  := 0,      // 未使能：设定冻结 / Idle, setpoint frozen
    eRun   := 10,     // 寻优运行中 / Optimisation active
    eFault := 90      // 故障锁存相（设定冻结保持） / Fault latched, setpoint frozen
);
END_TYPE

TYPE E_DL_VprCause :
(
    eNone       := 0, // 无故障成因 / No cause
    eCfgIllegal := 1, // 组态非法 / Illegal configuration
    eNonFinite  := 2  // 输入非有限 / Non-finite input
);
END_TYPE

FUNCTION_BLOCK FB_DL_VavPressureReset
VAR_INPUT
    fWorstDamperPct : REAL := 0.0;     // 最不利末端阀位 [%]，0~100 / Worst-case terminal damper position
    fDamperTargetPct: REAL := 90.0;    // 目标阀位 [%]，开区间 (0,100) / Target damper position
    fDeadbandPct    : REAL := 5.0;     // 阀位死区 [%]，域 >= 0 / Damper deadband
    fStepKpa        : REAL := 2.0;     // 单周期静压步长 [kPa]，域 > 0 / Static pressure step
    fSpMinKpa       : REAL := 100.0;   // 静压设定下限 [kPa] / Setpoint low limit
    fSpMaxKpa       : REAL := 500.0;   // 静压设定上限 [kPa] / Setpoint high limit
    fSpInitKpa      : REAL := 250.0;   // 设定初值（使能沿装载） [kPa] / Initial setpoint
    bEnable         : BOOL := FALSE;   // 寻优使能（电平）[-] / Optimisation enable
    bReset          : BOOL := FALSE;   // 复位命令，上升沿清故障 [-] / Reset edge
END_VAR
VAR_OUTPUT
    eState          : E_DL_VprState;   // 状态出口，段 6 单点映射 / State outlet
    eCause          : E_DL_VprCause;   // 故障成因出口（R190） / Fault cause outlet
    fSpKpa          : REAL;            // 静压设定输出 [kPa] / Static pressure setpoint
    bRaise          : BOOL;            // 本周期升压动作镜像 [-] / Raise action mirror
    bLower          : BOOL;            // 本周期降压动作镜像 [-] / Lower action mirror
    bError          : BOOL;            // 故障锁存标志 [-] / Fault latch flag
    nErrId          : UDINT;           // 故障码，0 = 无故障（本件无信息码） / Fault code only
END_VAR
VAR
    _eState         : E_DL_VprState := E_DL_VprState.eIdle;   // 内部相位（CASE 唯一写入目标） / Internal phase
    _eCause         : E_DL_VprCause := E_DL_VprCause.eNone;   // 故障成因锁存（锁存量） / Latched cause
    rtEnable        : R_TRIG;          // 使能沿实例，每周期无条件调用 / Enable edge
    rtReset         : R_TRIG;          // 复位沿实例，每周期无条件调用 / Reset edge
    _fSp            : REAL;            // 设定保持槽（持久） / Setpoint holding slot
    _fErrPct        : REAL;            // 阀位偏差 [%]（当拍量） / Damper deviation
    _bRaiseOn       : BOOL;            // 升压当拍量 [-] / Raise action
    _bLowerOn       : BOOL;            // 降压当拍量 [-] / Lower action
    _bNonFin        : BOOL;            // 输入非有限当拍量 [-] / Non-finite input
    _bCfgBad        : BOOL;            // 组态非法当拍量 [-] / Config illegal
    _bFault         : BOOL;            // 故障锁存位（锁存量） / Latched fault bit
    _uFault         : UDINT;           // 故障码锁存（锁存量） / Latched fault code
END_VAR

(* —— 段 0：沿实例无条件周期刷新 + 当拍量判据 —— *)
_fErrPct := fDamperTargetPct - fWorstDamperPct;                              // 阀位偏差 [%] / Damper deviation
_bNonFin := (fWorstDamperPct <> fWorstDamperPct) OR (fSpMinKpa <> fSpMinKpa)
         OR ((fWorstDamperPct - fWorstDamperPct) <> (fWorstDamperPct - fWorstDamperPct))
         OR ((fSpMinKpa - fSpMinKpa) <> (fSpMinKpa - fSpMinKpa));            // NaN 自反 + Inf 差值自减 / NaN and Inf
_bCfgBad := (fSpMaxKpa <= fSpMinKpa) OR (fStepKpa <= 0.0) OR (fDeadbandPct < 0.0)
            OR (fDamperTargetPct <= 0.0) OR (fDamperTargetPct >= 100.0);     // 组态非法当拍量 / Config illegal
rtEnable(CLK := bEnable);                                                    // 使能沿，每拍必调 / Enable edge
rtReset(CLK := bReset);                                                      // 复位沿，每拍必调 / Reset edge

(* —— 段 1：单拍量预清零（锁存量与设定保持槽不入清单） —— *)
bRaise := FALSE;                   // 升压镜像缺省 FALSE / Raise default
bLower := FALSE;                   // 降压镜像缺省 FALSE / Lower default
nErrId := 16#0000_0000;            // 故障码缺省无故障 / Fault code default

(* —— 段 2：复位沿 + 组态域闸 —— *)
IF rtReset.Q THEN                              // rtReset.Q = 当拍量 / current scan
    _bFault := FALSE;                          // 清故障锁存位（锁存量） / Clear fault latch
    _uFault := 16#0000_0000;                   // 清故障锁存码（锁存量） / Clear fault code
    _eCause := E_DL_VprCause.eNone;            // 清成因（锁存量） / Clear cause
    IF _eState = E_DL_VprState.eFault THEN
        _eState := E_DL_VprState.eIdle;        // 故障相迁出：回未使能 / Fault exit to idle
    END_IF
END_IF
IF _bCfgBad THEN                               // 组态域闸 / Config gate
    _uFault := 16#0002_0387;                   // 故障级：重置故障总码 / Algo fault code
    _eCause := E_DL_VprCause.eCfgIllegal;      // 归因：组态非法 / Cause: illegal config
    _bFault := TRUE;                           // 标志与码位配对（R45） / Flag paired with code
END_IF
IF (NOT _bFault) AND _bNonFin THEN             // 非有限锁存 / Non-finite latch
    _uFault := 16#0002_0387;
    _eCause := E_DL_VprCause.eNonFinite;       // 归因：非有限 / Cause: non-finite
    _bFault := TRUE;
END_IF

(* —— 段 3：寻优动作（仅在运行相且无故障；死区优先于动作） —— *)
IF (NOT _bFault) AND (_eState = E_DL_VprState.eRun) THEN
    IF ABS(_fErrPct) <= fDeadbandPct THEN                 // 死区内保持（容差式） / Deadband hold
        ;                                                // 保持：不动作 / Hold, no action
    ELSIF _fErrPct > fDeadbandPct THEN                    // 阀位偏小：升压 / Damper small: raise
        _fSp := _fSp + fStepKpa;                          // 单周期升压一个步长 / Raise one step
        _bRaiseOn := TRUE;
    ELSE                                                  // 阀位偏大：降压 / Damper large: lower
        _fSp := _fSp - fStepKpa;                          // 单周期降压一个步长 / Lower one step
        _bLowerOn := TRUE;
    END_IF
    IF _fSp < fSpMinKpa THEN                              // 下限钳制 / Low clamp
        _fSp := fSpMinKpa;
    ELSIF _fSp > fSpMaxKpa THEN                           // 上限钳制 / High clamp
        _fSp := fSpMaxKpa;
    END_IF
END_IF

(* —— 段 4：故障解除式（R240；全当拍量）：rtReset.Q / NOT _bCfgBad / NOT _bNonFin —— *)
IF rtReset.Q AND (NOT _bCfgBad) AND (NOT _bNonFin) THEN
    _bFault := FALSE;                          // 清故障锁存位（锁存量） / Clear fault latch
    _uFault := 16#0000_0000;                   // 清故障锁存码（锁存量） / Clear fault code
    _eCause := E_DL_VprCause.eNone;            // 清成因（锁存量） / Clear cause
END_IF

(* —— 段 4A：故障锁存相位迁移闸（设定冻结保持） —— *)
IF _bFault AND (_eState <> E_DL_VprState.eFault) THEN
    _eState := E_DL_VprState.eFault;           // 锁存即入故障相 / Latch enters fault phase
END_IF

(* —— 段 5：相位机（CASE 全覆盖 + ELSE 兜底） —— *)
CASE _eState OF

E_DL_VprState.eIdle:
    IF rtEnable.Q AND (NOT _bFault) THEN       // 使能上升沿：装载初值并钳制 / Enable edge loads initial value
        _fSp := fSpInitKpa;                    // 装载初值 / Load initial setpoint
        IF _fSp < fSpMinKpa THEN               // 初值下限钳制 / Initial low clamp
            _fSp := fSpMinKpa;
        ELSIF _fSp > fSpMaxKpa THEN            // 初值上限钳制 / Initial high clamp
            _fSp := fSpMaxKpa;
        END_IF
        _eState := E_DL_VprState.eRun;         // 进运行相 / Enter run
    END_IF

E_DL_VprState.eRun:
    IF NOT bEnable THEN                        // 撤使能：设定冻结，回未使能 / Disable: freeze and idle
        _eState := E_DL_VprState.eIdle;
    END_IF

E_DL_VprState.eFault:
    ;                                          // 故障相：设定冻结保持，仅段 4 复位沿可迁出 / Frozen, reset only

ELSE
    _uFault := 16#0002_0387;                   // 故障级：非法相位兜底（归并总码） / Illegal phase fallback
    _eCause := E_DL_VprCause.eCfgIllegal;      // 归因：相位非法归并组态 / Cause: phase illegal
    _bFault := TRUE;
    _eState := E_DL_VprState.eFault;           // 强制回故障相 / Force fault phase

END_CASE

(* —— 段 6：出口单点映射（名实同源；锁存码回放） —— *)
fSpKpa := _fSp;                                // 设定值出口 / Setpoint outlet
IF _bFault THEN
    nErrId := _uFault;                         // 故障锁存码回放 / Replay latched code
    bRaise := FALSE;                           // 故障相动作镜像强制 FALSE / Raise forced false
    bLower := FALSE;                           // 故障相动作镜像强制 FALSE / Lower forced false
ELSE
    nErrId := 16#0000_0000;                    // 无故障：本件无信息码 / No fault, no info code
    bRaise := _bRaiseOn;                       // 升压镜像 / Raise mirror
    bLower := _bLowerOn;                       // 降压镜像 / Lower mirror
END_IF
bError := _bFault;                             // 故障标志同源 / Flag from latch
eState := _eState;                             // 状态出口 / State outlet
eCause := _eCause;                             // 成因出口 / Cause outlet

END_FUNCTION_BLOCK

(* ---- FB_DL_AdaptiveLmsFilter.st ---- *)
(*
  ==================================================================
  组件名 Component  : FB_DL_AdaptiveLmsFilter
  分类   Category   : DL_Algo
  前缀   Naming     : FB_DL_ ｜ b/n/u/f/t/e/st 类型前缀制（R265）
  码位   Code ID    : 16#0002_374C（故障级）｜ 16#0002_3749 / 374A / 374B（信息级）
  版本   Version    : 1.0.1
  复杂度 Complexity  : 高
  功能   Purpose    : LMS 自适应横向滤波器（N 抽头权重在线更新 w[k] += 2μ·e·x[k]），
                      周期干扰对消 / 主动降噪的现场可整定基元。
  开源溯源 Origin    : 公开公式 clean-room，参考公开自适应信号处理教材的 LMS 权重
                      递推式（分类与公式借鉴，零代码复制），本件实现、闸门与码位
                      100% 自有。
  许可证 License    : MIT
  参考   Reference  : IEC 61131-3:2013 §6.6 算术运算符；LMS 递推 w[k] += 2μ·e·x[k]
                      为公开自适应滤波公式（Widrow-Hoff 类公开定义）
  平台   Platform   : 纯 IEC 61131-3（FOR / 四则 / R_TRIG / 比较），三平台通用
  依赖   Depends    : 仅 Standard.library（R_TRIG 属标准边沿检测）
  分工声明 Split     : FB_DL_BiquadFilter / FB_DL_BiquadCascade 为固定系数族；
                      FB_DL_DisturbanceObserver 为观测器路线；本件为在线自适应族；
                      互引 + MANUAL 选型段（「系数已知用 Biquad、干扰特征未知用
                      LMS」）（R216）。
  归属 Ownership     : 本件无 TYPE 声明；全部引脚为 IEC 标准原生类型。
  ------------------------------------------------------------------
  边界 Boundary     :
                      一 延迟线固定 ARRAY[0..31] OF LREAL（禁动态分配），每拍右移
                         入 fRef；uTaps 越域钳位 4..32 + 信息级 374A，钳位赋值
                         上移至变更沿检测前（R64 v1.0.1）：抽头数变更沿以本拍
                         钳位值判定，无晚一拍混算窗口（旧值配新权重 / 延迟线
                         的混算拍已消除）；变更沿清权重与延迟线（活动抽头数才
                         参与运算）；
                      二 fMu 域闸 (0, 0.1] 且非有限 → 组态码 3749 + 权重冻结 +
                         三件套 + RETURN 结构早退；
                      三 任一输入非有限（fRef / fDesired）→ 权重冻结 + 故障码 374C
                         + bValid = FALSE；两条恢复路径拆明（R64 v1.0.1）：
                         a) NaN 输入（测点坏）——权重未被写入污染物，测点恢复后
                            下一拍自动恢复；b) 溢出污染——权重写回前 |corr·x|
                            预检命中非有限即 374C 冻结（跳过写回），若上一拍已
                            写入污染物则需 bWipeW 才能恢复（不可自动恢复性写死）；
                         递推结果复检非有限同码处置（更新前置闸：命中路径冻结
                         权重，禁污染物写入）；
                      四 fWEnergy > 1.0E12 → 发散监视信息级 374B（建议减小 μ，不
                         自动清权重，诊断出口，每拍重算不锁存）；374B 为持续
                         发散监视，溢出（写回预检命中）当拍改报故障级 374C 并
                         早退，溢出一次性报告、374B 不逐拍重报溢出
                         （R64 v1.0.1 口径）；
                      五 bWipeW 单拍 → 全权重与延迟线清零（段 0 R_TRIG 无条件刷新）；
                      六 bEnable = FALSE 的语义写死（FB33-4 声明行）：权重保留但
                         停止更新、fErr 冻结——现场断使能调试时不丢已收敛权重；
                      七 故障码策略（本件无 bReset 引脚，R152 解除路径自证）：组态
                         与测量类故障码逐拍重算不锁存，解除路径 = 修正组态 / 测点
                         恢复（恒可达）；发散信息级逐拍重算；
                      八 段 0 无条件刷新 R_TRIG；CASE 无（线性递推，R6 标注 N/A）；
                         首拍 _bInit 全量初始化；无全局、无外部变量、无物理地址。
  错误码 Codes      :
    16#0002_3749【故障级】组态非法（fMu ≤ 0 / > 0.1 / 非有限）
    16#0002_374A【信息级】uTaps 越域已钳位（合法 4..32，不置 bError）
    16#0002_374B【信息级】权重平方和超阈（fWEnergy > 1.0E12，持续发散监视，建议
                         减小 μ；溢出当拍由 374C 承担并早退，374B 不重报溢出）
    16#0002_374C【故障级】输入非有限（fRef / fDesired 为 NaN / ±Inf）、递推结果
                         非有限、或权重写回前 |corr·x| 预检命中非有限（溢出污染，
                         需 bWipeW 恢复，出口同形 R90）
  码位反证 Note     :
    3749 与 374C 不可合并：3749 与输入无关（组态即刻判），374C 需输入到达，处置人
    不同（组态工程师 / 现场测点），可由场景还原（R90）；374A / 374B 信息级子带
    （R75 纪律），不跨用故障子带。
  验收 Acceptance   :
    算法已证（脚本）：未跑 ｜ 编译器已证（三平台）：未跑
    V1 fRef = 0 → 权重不增长、fErr = fDesired
    V2 正弦干扰 + 相关参考 → fErr 包络逐拍递减（定性收敛向量）
    V3 fMu = 0 → 组态早退权重冻结；V4 fRef = NaN 单拍 → 权重冻结 + 故障
       （下一拍恢复后 fErr 不含污染：权重未变断言）
    V5 uTaps = 100 → 钳 32 + 信息级；V6 bWipeW → fWEnergy = 0
    V7 权重平方和超阈 → 信息级不锁存
  修订记录 Revision  :
    2026-11-21  v1.0.0  R63 首版（批 4 · 序号 11）
    2026-11-21  v1.0.1  R64 返修 R63-D3/D4：抽头数钳位赋值整体上移至段 4 变更沿
                        检测前（变更沿以本拍钳位值判定，无晚一拍混算窗口）；
                        段 11 写回前 ABS(_fCorr*_afX[_i]) 预检，命中即 374C 冻结
                        权重当拍早退（溢出一次性报告），374B 改持续发散监视；
                        边界三拆明两条恢复路径（NaN 输入自动恢复 / 溢出需
                        bWipeW），删除「理论上不可达」失准表述
  ==================================================================
*)
FUNCTION_BLOCK FB_DL_AdaptiveLmsFilter
VAR_INPUT
    bEnable   : BOOL := TRUE;   // 使能，FALSE 时权重保留但停止更新（边界六）/ the enable, false keeps the weights but stops the update
    bWipeW    : BOOL := FALSE;  // 权重清零电平，上升沿全权重与延迟线清零 / the wipe level, its rising edge clears the weights and the delay line
    fRef      : LREAL := 0.0;   // 参考输入 [工程单位]（与干扰相关的信号）/ the reference input correlated with the disturbance
    fDesired  : LREAL := 0.0;   // 主输入 [工程单位] / the desired main input
    uTaps     : USINT := 16;    // 抽头数 [个]，合法域 4..32，变更沿清权重 / the tap count, legal four to thirty two
    fMu       : LREAL := 0.01;  // 步长 [−]，域 (0, 0.1] / the step size inside the half open domain
END_VAR
VAR_OUTPUT
    fErr      : LREAL := 0.0;           // 误差 = fDesired − fOut [工程单位] / the error of the desired minus the output
    fOut      : LREAL := 0.0;           // 滤波输出 [工程单位] / the filter output
    fWEnergy  : LREAL := 0.0;           // 权重平方和 [−]，收敛 / 发散诊断 / the squared weight sum for the convergence diagnostics
    bValid    : BOOL := FALSE;          // 输出可用 [-] / the output is usable
    eErr      : UDINT := 16#0000_0000;  // 错误码，0 = 正常 / the error code, zero is ok
    bError    : BOOL := FALSE;          // 故障标志（故障级码同拍置位，R45 配对）/ the fault flag raised with a fault level code
END_VAR
VAR
    _bInit    : BOOL := FALSE;              // 首拍初始化标志（R310 / FB50-2）/ the first scan flag
    _afW      : ARRAY[0..31] OF LREAL;      // 权重数组 [−]，固定 32 抽头 / the fixed weight array of thirty two taps
    _afX      : ARRAY[0..31] OF LREAL;      // 延迟线 [工程单位] / the delay line
    _nTaps    : DINT := 16;                 // 钳位后的抽头数 [个] / the clamped tap count
    _nTapsPrev: DINT := 0;                  // 上拍抽头数快照 [个]，置 0 使首拍必触发清权重 / the previous tap count
    _i        : DINT := 0;                  // 抽头遍历索引 [下标] / the tap traversal index
    _iShift   : DINT := 0;                  // 移位遍历索引 [下标] / the shift traversal index
    _fAcc     : LREAL := 0.0;               // 输出累加器 [工程单位] / the output accumulator
    _fEng     : LREAL := 0.0;               // 权重能量累加器 [−] / the weight energy accumulator
    _fErrUse  : LREAL := 0.0;               // 误差工作副本 [工程单位] / the working error copy
    _fCorr    : LREAL := 0.0;               // 修正量 2μ·e [−] / the correction factor of two mu times the error
    _fProdAbs : LREAL := 0.0;               // 写回预检量 |corr·x| [−]（R64 v1.0.1）/ the writeback precheck magnitude of the correction times the tap
    _bWOverflow: BOOL := FALSE;             // 写回预检溢出命中标记（单拍，R64 v1.0.1）/ the writeback overflow hit flag of this scan
    _bFinRef  : BOOL := FALSE;              // 参考输入有限闸结果（逐拍重算）/ the reference finiteness gate result
    _bFinDes  : BOOL := FALSE;              // 主输入有限闸结果（逐拍重算）/ the desired finiteness gate result
    _bFinMu   : BOOL := FALSE;              // 步长有限闸结果（逐拍重算）/ the mu finiteness gate result
    _bCfgBad  : BOOL := FALSE;              // 组态非法标记（逐拍重算）/ the configuration fault flag
    _bTapClamp: BOOL := FALSE;              // 抽头数钳位标记（逐拍重算，信息级 374A）/ the tap clamp flag
    _bDivWarn : BOOL := FALSE;              // 发散警告标记（逐拍重算，信息级 374B）/ the divergence warning flag
    rtWipe    : R_TRIG;                     // 权重清零沿实例，段 0 无条件刷新（R7）/ the wipe edge instance refreshed unconditionally
END_VAR  // R64 结构补齐：VAR 段缺失的 END_VAR（门禁机械修复）
VAR CONSTANT
    DL_LMS_TMAX  : DINT := 32;        // 抽头容量上界 [个]，与数组容量一致 / the tap capacity aligned with the array
    DL_LMS_TMIN  : DINT := 4;         // 抽头数下界 [个] / the tap floor
    DL_LMS_MUMAX : LREAL := 0.1;      // 步长上界 [−] / the step size ceiling
    DL_LMS_MUZERO: LREAL := 0.0;      // 步长零常量 [−] / the step size zero constant
    DL_LMS_TWO   : LREAL := 2.0;      // LMS 修正系数常量 [−] / the LMS correction factor constant
    DL_LMS_WMAX  : LREAL := 1.0E12;   // 权重平方和发散门限 [−] / the divergence threshold of the weight energy
    DL_LMS_ZERO  : LREAL := 0.0;      // 实数零常量 [工程单位] / the real zero constant
    DL_LMS_ZEROI : DINT := 0;         // 整型零常量 [个] / the integer zero constant
    DL_LMS_ONEI  : DINT := 1;         // 整型一常量 [个] / the integer one constant
END_VAR

// 段 0｜组态闸先行 + 沿检测无条件周期刷新（禁入分支，R7）/ segment 0, the configuration gate first and the unconditional edge refresh
_bFinMu := (fMu = fMu) AND ((fMu - fMu) = (fMu - fMu)); // 步长有限 / the step size is finite
_bCfgBad := (NOT _bFinMu) OR (fMu <= DL_LMS_MUZERO) OR (fMu > DL_LMS_MUMAX); // 组态非法 / an illegal configuration
rtWipe(CLK := bWipeW); // 权重清零沿 / the wipe edge

// 段 1｜首拍初始化（FB50-2）/ segment 1, the first scan init
IF NOT _bInit THEN // 首拍一拍 / the first scan
    _bInit := TRUE; // 置首拍标志 / raise the first scan flag
    _nTapsPrev := DL_LMS_ZEROI; // 抽头数快照置 0，使段 4 变更沿必然触发一次清权重 / zero the snapshot so the change edge clears the weights once
    FOR _i := DL_LMS_ZEROI TO DL_LMS_TMAX - DL_LMS_ONEI DO // 有界遍历全容量 / the bounded traversal over the full capacity
        _afW[_i] := DL_LMS_ZERO; // 权重显式清零 [−] / clear the weight explicitly
        _afX[_i] := DL_LMS_ZERO; // 延迟线显式清零 [工程单位] / clear the delay line explicitly
    END_FOR
END_IF

// 段 2｜单拍量预置 / segment 2, the per scan preset
_bTapClamp := FALSE; // 钳位标记预清零（单拍信息位，段 7 映射）/ preset the clamp flag false
_bDivWarn := FALSE; // 发散警告标记预清零（单拍信息位）/ preset the divergence flag false
_fErrUse := fErr; // 误差工作副本接管上拍出口（冻结语义基线）[工程单位] / the working error takes the previous outlet as the freeze base

// 段 3｜组态非法结构早退：权重冻结（边界二，出口三件套 + RETURN）/ segment 3, the structural early exit on an illegal configuration
IF _bCfgBad THEN // 组态非法 / an illegal configuration
    bValid := FALSE; // 输出不可用 / the output is not usable
    eErr := 16#0002_3749; // 故障级：组态非法 / fault grade, an illegal configuration
    bError := TRUE; // 同拍置故障标志（R45 配对）/ raise the fault flag on the same scan
    RETURN; // 结构早退，权重冻结（禁污染）/ the structural early exit with the weights frozen
END_IF

// 段 4｜抽头数钳位（边界一，信息级 374A；R64 v1.0.1 整体上移至变更沿检测前，
//        保证段 5 变更沿以本拍钳位值判定，无晚一拍混算窗口）/ segment 4, the tap clamp moved before the change edge
_nTaps := USINT_TO_DINT(uTaps); // 抽头数升位接管 [个] / take the tap count widened
IF (_nTaps < DL_LMS_TMIN) OR (_nTaps > DL_LMS_TMAX) THEN // 抽头数越域 / the count is out of the domain
    _bTapClamp := TRUE; // 置钳位标记（信息级 374A）/ raise the clamp flag
    IF _nTaps < DL_LMS_TMIN THEN // 下界钳位 / the floor clamp
        _nTaps := DL_LMS_TMIN; // 钳到下界 [个] / clamp to the floor
    ELSE // 上界钳位 / the ceiling clamp
        _nTaps := DL_LMS_TMAX; // 钳到容量 [个] / clamp to the capacity
    END_IF
END_IF

// 段 5｜权重清零沿：全权重与延迟线清零（边界五；抽头数变更沿同段处理，
//        以段 4 本拍钳位值判定）/ segment 5, the wipe edge and the tap change edge
IF (_nTaps <> _nTapsPrev) OR rtWipe.Q THEN // 抽头数变更沿或清零沿 / the tap change edge or the wipe edge
    FOR _i := DL_LMS_ZEROI TO DL_LMS_TMAX - DL_LMS_ONEI DO // 有界遍历全容量 / the bounded traversal over the full capacity
        _afW[_i] := DL_LMS_ZERO; // 权重清零 [−] / clear the weight
        _afX[_i] := DL_LMS_ZERO; // 延迟线清零 [工程单位] / clear the delay line
    END_FOR
    _nTapsPrev := _nTaps; // 快照本拍抽头数 / snapshot the tap count
END_IF

// 段 6｜失能分支：权重保留但停止更新（边界六声明行）/ segment 6, the disabled branch keeps the weights
IF NOT bEnable THEN // 失能 / disabled
    bValid := FALSE; // 输出不可用 / the output is not usable while disabled
    bError := FALSE; // 失能不是故障 / a disabled device is not a fault
    eErr := 16#0000_0000; // 失能不发码 / no code is emitted while disabled
    RETURN; // 早退，权重保留（现场断使能调试不丢已收敛权重）/ early return with the weights kept
END_IF

// 段 7｜输入非有限闸：权重冻结（边界三，禁污染权重）/ segment 7, the input finiteness gate freezes the weights
_bFinRef := (fRef = fRef) AND ((fRef - fRef) = (fRef - fRef)); // 参考输入有限 / the reference is finite
_bFinDes := (fDesired = fDesired) AND ((fDesired - fDesired) = (fDesired - fDesired)); // 主输入有限 / the desired is finite
IF (NOT _bFinRef) OR (NOT _bFinDes) THEN // 任一输入坏 / either input is broken
    bValid := FALSE; // 输出不可用 / the output is not usable
    eErr := 16#0002_374C; // 故障级：输入非有限 / fault grade, an input is not finite
    bError := TRUE; // 同拍置故障标志（R45 配对）/ raise the fault flag on the same scan
    RETURN; // 早退，权重冻结（不更新，污染不可自动恢复性见边界三）/ early return with the weights frozen
END_IF

// 段 8｜延迟线右移入新样本（边界一，固定容量，禁动态分配）/ segment 8, the delay line shifts the new sample in
FOR _iShift := DL_LMS_TMAX - DL_LMS_ONEI TO DL_LMS_ONEI BY -1 DO // 有界逆向遍历（31 → 1）/ the bounded reverse traversal from thirty one down to one
    _afX[_iShift] := _afX[_iShift - DL_LMS_ONEI]; // 延迟线逐位右移 [工程单位] / shift the delay line one slot right
END_FOR
_afX[DL_LMS_ZEROI] := fRef; // 新样本入延迟线首槽 [工程单位] / the new sample enters the first slot

// 段 9｜滤波输出与误差计算（活动抽头数才参与，边界一）/ segment 9, the output and the error over the active taps
_fAcc := DL_LMS_ZERO; // 输出累加器清零 [工程单位] / clear the output accumulator
FOR _i := DL_LMS_ZEROI TO _nTaps - DL_LMS_ONEI DO // 有界遍历活动抽头（上界已证 ≤ 32）/ the bounded traversal over the active taps
    _fAcc := _fAcc + (_afW[_i] * _afX[_i]); // 横向滤波加权和 [工程单位] / the transversal weighted sum
END_FOR
fOut := _fAcc; // 滤波输出出口 [工程单位] / the filter output outlet
_fErrUse := fDesired - fOut; // 误差 = 主输入 − 输出 [工程单位] / the error of the desired minus the output

// 段 10｜递推结果复检（更新前置闸：结果非有限则权重冻结，禁污染物写入，边界三）/ segment 10, the result recheck before the update
IF (_fErrUse <> _fErrUse) OR ((_fErrUse - _fErrUse) <> (_fErrUse - _fErrUse))
OR (fOut <> fOut) OR ((fOut - fOut) <> (fOut - fOut)) THEN // 误差或输出非有限（理论上不可达，防御保留）/ a non finite error or output
    bValid := FALSE; // 输出不可用 / the output is not usable
    eErr := 16#0002_374C; // 故障级：输入或结果非有限（同族一码，出口同形，R90）/ fault grade under the same family code
    bError := TRUE; // 同拍置故障标志（R45 配对）/ raise the fault flag on the same scan
    RETURN; // 早退，权重冻结 / early return with the weights frozen
END_IF

// 段 11｜LMS 权重在线更新（公开公式：w[k] += 2μ·e·x[k]，边界三判据已过）；
//         写回前 |corr·x| 预检（R64 v1.0.1，R63-D4）：命中非有限即 374C 冻结
//         权重当拍早退（跳过写回与段 12 的 374B 判定，溢出一次性报告）/
//         segment 11, the LMS weight update with the writeback precheck
_fCorr := DL_LMS_TWO * fMu * _fErrUse; // 修正量 2μ·e [−] / the correction factor
_bWOverflow := FALSE; // 预检命中标记预清零（单拍量，本段内置）/ preset the overflow hit flag false
FOR _i := DL_LMS_ZEROI TO _nTaps - DL_LMS_ONEI DO // 有界遍历活动抽头 / the bounded traversal over the active taps
    _fProdAbs := ABS(_fCorr * _afX[_i]); // 写回预检量 |corr·x| [−]（先算后判，命中即冻结）/ the precheck magnitude computed before the writeback
    IF (_fProdAbs <> _fProdAbs) OR ((_fProdAbs - _fProdAbs) <> (_fProdAbs - _fProdAbs)) THEN // 预检量非有限（NaN 或 ±Inf，溢出真实可达：μ 上界 0.1 内大误差大样本即可触发）/ a non finite precheck magnitude, reachable on the overflow
        _bWOverflow := TRUE; // 置溢出命中标记 / raise the overflow hit flag
        EXIT; // 跳出写回（冻结权重，禁污染物写入）/ leave the loop without the writeback, the weights stay frozen
    END_IF
    _afW[_i] := _afW[_i] + (_fCorr * _afX[_i]); // 权重递推 [−]（预检已过才写回）/ the weight recursion only after the precheck passed
END_FOR
IF _bWOverflow THEN // 预检命中：溢出一次性报告（故障级 374C，本拍不进段 12 的 374B 判定，R64 v1.0.1）/ the precheck hit, the overflow is reported once
    fErr := _fErrUse; // 误差出口照实（已过段 10 有限闸）[工程单位] / the error outlet is still finite
    bValid := FALSE; // 输出不可用 / the output is not usable
    eErr := 16#0002_374C; // 故障级：写回预检命中非有限（溢出污染，需 bWipeW 恢复，边界三路径 b）/ fault grade, the writeback precheck hit a non finite magnitude
    bError := TRUE; // 同拍置故障标志（R45 配对）/ raise the fault flag on the same scan
    RETURN; // 早退，权重冻结（跳过段 12 能量诊断，374B 本拍不判）/ early return with the weights frozen, the energy diagnostics are skipped this scan
END_IF
fErr := _fErrUse; // 误差出口（已过有限闸）[工程单位] / the error outlet after the gate

// 段 12｜权重能量诊断（边界四，信息级 374B，每拍重算不锁存）/ segment 12, the weight energy diagnostics
_fEng := DL_LMS_ZERO; // 能量累加器清零 [−] / clear the energy accumulator
FOR _i := DL_LMS_ZEROI TO _nTaps - DL_LMS_ONEI DO // 有界遍历活动抽头 / the bounded traversal over the active taps
    _fEng := _fEng + (_afW[_i] * _afW[_i]); // 权重平方累加 [−] / accumulate the squared weights
END_FOR
fWEnergy := _fEng; // 权重平方和出口 [−] / the weight energy outlet
IF fWEnergy > DL_LMS_WMAX THEN // 超发散门限 / above the divergence threshold
    _bDivWarn := TRUE; // 置发散警告标记（信息级 374B）/ raise the divergence flag
END_IF

// 段 13｜统一出口（信息级重算，R187 / FB51-8）/ segment 13, the unified outlet
bValid := TRUE; // 输出可用 / the output is usable
bError := FALSE; // 无故障 / no fault
IF _bTapClamp THEN // 抽头数钳位（信息级，逐拍重算）/ the tap clamp, informational
    eErr := 16#0002_374A; // 信息级：uTaps 越域已钳位 / informational, the tap count was clamped
ELSIF _bDivWarn THEN // 发散警告（信息级，逐拍重算）/ the divergence, informational
    eErr := 16#0002_374B; // 信息级：权重平方和超阈，建议减小 μ / informational, the weight energy is over the threshold, reduce the step size
ELSE // 无事件 / no event
    eErr := 16#0000_0000; // 正常 / ok
END_IF
END_FUNCTION_BLOCK

(* ---- FB_DL_BiquadFilter.st ---- *)
(*
  ==================================================================
  组件名 Component  : FB_DL_BiquadFilter
  分类   Category   : DL_Algo
  前缀   Naming     : FB_DL_ ｜ b/n/u/f/t/e/st 类型前缀制（R265）
  码位   Code ID    : 16#0002_3735 / 3736 / 3737 / 373A（故障级）
                      16#0002_3738 / 3739（信息级）
  版本   Version    : 1.0.1
  复杂度 Complexity  : 高
  功能   Purpose    : 通用二阶 IIR 节（Direct Form I），系数由调用方下发（归一化 a0 = 1），
                      可配低通 / 高通 / 带通 / 带阻 / 全通；带 Jury 三条件稳定域闸、
                      系数变更沿清状态、输出钳位 + 抗 windup 状态回写。
  开源溯源 Origin    : IEC 61131-3 标准语义的道莅防御性实现（clean-room，无第三方代码行）；
                      差分方程与三角稳定判据取自公开 DSP 教科书与公开滤波器设计手册的
                      通用公式（分类与公式借鉴，零代码复制），本件实现、闸门与码位 100% 自有。
  许可证 License    : MIT
  参考   Reference  : IEC 61131-3:2013 §6.6 算术运算符；二阶 IIR 直接I型差分方程的公开
                      定义（RBJ Audio EQ Cookbook 类公开二阶节设计公式，仅借鉴公式结构）
  平台   Platform   : 纯 IEC 61131-3（四则 / ABS / R_TRIG / 比较），三平台通用
  依赖   Depends    : 仅 Standard.library（R_TRIG 属标准边沿检测）
  分工声明 Split     : FB_DL_LowPassFilter（一阶 RC）/ FB_DL_HighPassFilter（一阶）/
                      FB_DL_NotchFilter（陷波专用，结构固定）/ FB_DL_FirFilter（FIR）
                      为结构专用轻量件；本件为通用二阶节，适用于「需要带通 / 带阻 /
                      可调 Q 且带 ST 系数下发」的场合（R216 双向互引，选型对照见
                      MANUAL_DL_Algo）。
  归属 Ownership     : 本件无 TYPE 声明；全部引脚为 IEC 标准原生类型。
  ------------------------------------------------------------------
  边界 Boundary     :
                      一 稳定域闸（v1.0.1 返修 R63 · 修 R62-D2 严重：换 Jury 三条件，废除
                         「|a1|<2 且 |a2|<1 且 |a2−a1|<1」伪判据——该伪判据放行了
                         a1 = −1.9 / a2 = −0.95 的实根 −0.9545 发散极点族）：判据为
                         ABS(a2) < 1 且 (1 + a1 + a2) > 0 且 (1 − a1 + a2) > 0，
                         任一不满足即判组态故障并冻结输出，绝不外泄发散值；
                      二 系数任一非有限（NaN / ±Inf）同走组态故障路径；八个浮点入参
                         （fIn / b0 / b1 / b2 / a1 / a2 / fOutMin / fOutMax）逐个点名闸，
                         换算量与限值一并入闸（R272，禁按「主要参数」手挑）；
                      三 系数变更沿（五系数任一 |新 − 旧| > 1.0E-9）清 w1 / w2：防旧状态
                         冲击新频响，属「在线变系数为无扰切换的保守处置」，非无扰切换本身；
                      四 输出钳位 + 抗 windup：fOut 钳 [fOutMin, fOutMax]，被钳时 w1 := fOut
                         回写状态，防积分式累积发散；
                      五 bEnable = FALSE 的语义二选一并写死（FB33-4 声明行）：本件取
                         「降级为安全值 0.0 + 状态清零 + bValid = FALSE」，理由：滤波器输出
                         是下游控制量，失能须归零而非冻结末值；
                      六 故障码一律锁存至 bResetState 上升沿回放，不在故障相按当下输入
                         重新推断（FB33-1 / R152：首因不会被末因覆盖）；清除路径 = 复位沿；
                      七 信息级码（输出钳位 / 系数变更）逐拍重算不锁存；
                      八 段 0 无条件刷新 R_TRIG；CASE 无（本件为线性节，无顺序状态机，
                         R6 标注 N/A），故 ELSE 兜底要求不适用；首拍 _bInit 初始化全量状态。
  错误码 Codes      :
    16#0002_3735【故障级】系数越过 Jury 三条件稳定域（|a2| ≥ 1 或 1+a1+a2 ≤ 0 或
                         1−a1+a2 ≤ 0），锁存
    16#0002_3736【故障级】系数非有限（五个系数任一为 NaN 或 ±Inf），锁存
    16#0002_3737【故障级】输出钳位域非法（fOutMin > fOutMax 或限值非有限），锁存
    16#0002_3738【信息级】本拍输出被钳位（bSat = TRUE，不锁存）
    16#0002_3739【信息级】系数变更沿触发状态清零（不锁存）
    16#0002_373A【故障级】输入 / 中间量 / 输出非有限（NaN 或 ±Inf），锁存；
                         v1.0.1 返修（R63 · 修 R62-D5）：本码路径不再复用 bCfgBad 表达，
                         改由 bValid = FALSE + eErr = 373A 单独承载（bCfgBad 专指组态族）
  码位反证 Note     :
    3735 / 3736 / 3737 / 373A 四码不可合并：四者的 bCfgBad 与 bValid 组合完全相同，
    现场若只靠输出组合无法区分「系数发散 / 系数采集失败 / 限值配错 / 输入测点坏」，
    而四者的处置人不同（算法工程师 / 仪表工 / 组态工程师 / 现场仪表）（R90 反证句）。
  验收 Acceptance   :
    算法已证（脚本）：未跑 ｜ 编译器已证（三平台）：未跑
    V1 阶跃输入 + 公开二阶低通系数组（b0 = 0.0675, b1 = 0.1349, b2 = 0.0675,
       a1 = -1.1430, a2 = 0.4128）→ 输出单调收敛于稳态 1.0，无过冲爆炸（极点半径 √0.4128 ≈ 0.6426）
    V2 a1 = 2.5（不稳定）→ bCfgBad = TRUE + fOut 冻结 + 码 3735
    V2b a1 = -1.9, a2 = -0.95（v1.0.1 返修向量：旧伪判据放行的发散族）→ Jury 判
       3735 + fOut 冻结 + bCfgBad = TRUE（ABS(a2)=0.95 < 1 成立但 1+a1+a2 = -1.85 ≤ 0 不满足）
    V2c a1 = 0.0, a2 = -0.99（v1.0.1 返修向量：合法边界内）→ Jury 三条件全成立，
       合法放行（旧 |a2−a1|<1 伪判据对该族误杀）
    V3 a1 = NaN → 同 V2，码 3736
    V4 在线把低通系数换成高通系数 → w1 / w2 清零，fOut 单拍跳变被钳位而不发散，码 3739
    V5 bResetState 单拍 → w1 = w2 = 0
    V6 fIn = 1.0E9 持续 → fOut 钳 fOutMax + bSat + w1 回写（下一拍不反向冲）
    V7 bEnable = FALSE → fOut = 0.0、状态零、bValid = FALSE
    V8 fOutMin > fOutMax → 码 3737 + bCfgBad
    V9 首拍 → 状态零、fOut = 0.0（禁首拍用未初始化状态）
  修订记录 Revision  :
    2026-11-21  v1.0.0  R62 首版（批 3 · 序号 9）
    2026-11-21  v1.0.1  R63 返修 R2（R62-D2 严重 + D5 轻）：①稳定判据换 Jury 三条件
                        ABS(a2)<1 ∧ (1+a1+a2)>0 ∧ (1−a1+a2)>0，码 3735 语义与头注释同步；
                        ②新增验收向量 V2b（旧伪判据放行族判 3735+冻结）与 V2c（合法边界族放行）；
                        ③373A（输入/中间/输出非有限）路径不再复用 bCfgBad，改 bValid+eErr 表达
  ==================================================================
*)
FUNCTION_BLOCK FB_DL_BiquadFilter
VAR_INPUT
    bEnable     : BOOL := TRUE;    // 使能；FALSE 时输出归零并清状态（边界五）/ the enable, false zeroes the output and clears the state
    bResetState : BOOL := FALSE;   // 状态复位电平，上升沿清 w1 / w2 与故障锁存 / the state reset level, its rising edge clears the states and the fault latch
    fIn         : LREAL := 0.0;    // 输入量 [工程单位]，必须有限 / the input value, must be finite
    fB0         : LREAL := 1.0;    // 归一化前向系数 b0 [−]，a0 已归一为 1 / the normalized feed forward coefficient b0
    fB1         : LREAL := 0.0;    // 归一化前向系数 b1 [−] / the normalized feed forward coefficient b1
    fB2         : LREAL := 0.0;    // 归一化前向系数 b2 [−] / the normalized feed forward coefficient b2
    fA1         : LREAL := 0.0;    // 归一化反馈系数 a1 [−]，须落三角稳定域 / the normalized feedback coefficient a1 inside the triangle
    fA2         : LREAL := 0.0;    // 归一化反馈系数 a2 [−]，须落三角稳定域 / the normalized feedback coefficient a2 inside the triangle
    fOutMin     : LREAL := -1.0E6; // 输出钳位域下界 [工程单位] / the output clamp floor
    fOutMax     : LREAL := 1.0E6;  // 输出钳位域上界 [工程单位] / the output clamp ceiling
    tSample     : TIME := T#10MS;  // 采样周期 [毫秒]，仅作标称记录（系数设计已内含采样率）/ the nominal sample period, recorded only
END_VAR
VAR_OUTPUT
    fOut    : LREAL := 0.0;           // 滤波输出 [工程单位] / the filtered output
    bSat    : BOOL := FALSE;          // 本拍输出被钳位 [-] / the output was clamped on this scan
    bCfgBad : BOOL := FALSE;          // 组态非法（与故障锁存同源，锁存型）[-] / an illegal configuration, latched with the fault
    bValid  : BOOL := FALSE;          // 输出可用（失能 / 故障 / 输入非有限为 FALSE）[-] / the output is usable
    eErr    : UDINT := 16#0000_0000;  // 错误码，0 = 正常 / the error code, zero is ok
    bError  : BOOL := FALSE;          // 故障锁存位（由锁存码派生，非单拍标志，R99）/ the latched fault bit derived from the latched code
END_VAR
VAR
    _bInit     : BOOL := FALSE;               // 首拍初始化标志（R310 / FB50-2）/ the first scan flag
    _fW1       : LREAL := 0.0;                // 状态 w1（上一拍中间量）[工程单位] / the state w1 of the previous scan
    _fW2       : LREAL := 0.0;                // 状态 w2（前两拍中间量）[工程单位] / the state w2 of two scans ago
    _fW        : LREAL := 0.0;                // 本拍中间量 w [工程单位] / the intermediate w of this scan
    _fY        : LREAL := 0.0;                // 本拍未钳位输出 y [工程单位] / the unclamped output y of this scan
    _fOutLast  : LREAL := 0.0;                // 最近一次有效输出（故障冻结源）[工程单位] / the last valid output used while frozen
    _fB0Prev   : LREAL := 0.0;                // 上拍 b0 快照 [−] / the previous b0 snapshot
    _fB1Prev   : LREAL := 0.0;                // 上拍 b1 快照 [−] / the previous b1 snapshot
    _fB2Prev   : LREAL := 0.0;                // 上拍 b2 快照 [−] / the previous b2 snapshot
    _fA1Prev   : LREAL := 0.0;                // 上拍 a1 快照 [−] / the previous a1 snapshot
    _fA2Prev   : LREAL := 0.0;                // 上拍 a2 快照 [−] / the previous a2 snapshot
    _bFinCoef  : BOOL := FALSE;               // 五个系数有限闸结果（逐拍重算）/ the coefficient finiteness gate result
    _bFinIn    : BOOL := FALSE;               // 输入有限闸结果（逐拍重算）/ the input finiteness gate result
    _bFinDom   : BOOL := FALSE;               // 钳位域合法闸结果（逐拍重算）/ the clamp domain gate result
    _bStable   : BOOL := FALSE;               // Jury 三条件稳定域闸结果（逐拍重算，v1.0.1 换判据）/ the Jury three condition stability gate result
    _bCfgBadI  : BOOL := FALSE;               // 本拍组态非法标记（逐拍重算）/ the per scan configuration fault flag
    _bCoefChg  : BOOL := FALSE;               // 系数变更沿标记（逐拍重算，信息级 3739）/ the coefficient change flag
    _bSatI     : BOOL := FALSE;               // 本拍钳位内部位，段 1 预清段 12 映射 / the internal clamp bit
    _uLatch    : UDINT := 16#0000_0000;       // 故障码锁存（仅复位沿清除，FB33-1）/ the latched fault code cleared only by the reset edge
    rtReset    : R_TRIG;                      // 复位沿实例，段 0 无条件刷新（R7）/ the reset edge instance refreshed unconditionally
END_VAR  // R64 结构补齐：VAR 段缺失的 END_VAR（门禁机械修复）
VAR CONSTANT
    DL_BQ_EPS    : LREAL := 1.0E-9; // 系数变更判定容差 [−]，浮点禁判等 / the coefficient change tolerance, plain equality is forbidden
    DL_BQ_A2LIM  : LREAL := 1.0;    // Jury 条件一 |a2| 边界 [−] / the Jury first condition boundary on the absolute a2
    DL_BQ_ONE    : LREAL := 1.0;    // Jury 条件二三的一常量 [−] / the unit constant of the Jury second and third conditions
    DL_BQ_ZERO   : LREAL := 0.0;    // 实数零常量 [工程单位] / the real zero constant
END_VAR

// 段 0｜沿检测无条件周期刷新（禁入分支，R7）/ segment 0, the unconditional edge refresh
rtReset(CLK := bResetState); // 复位沿 / the reset edge

// 段 1｜首拍初始化与单拍标志预清（R310 / FB32-1；_bInit 与复位沿同款初始化）/ segment 1, the first scan init and the preset
IF NOT _bInit THEN // 首拍一拍 / the first scan
    _bInit := TRUE; // 置首拍标志 / raise the first scan flag
    _fW1 := DL_BQ_ZERO; // 状态 w1 显式清零 / clear the state w1 explicitly
    _fW2 := DL_BQ_ZERO; // 状态 w2 显式清零 / clear the state w2 explicitly
    _fOutLast := DL_BQ_ZERO; // 最近有效输出显式清零（禁首拍用未初始化状态）/ clear the last valid output explicitly
    _uLatch := 16#0000_0000; // 故障码锁存显式清零 / clear the latched code explicitly
    _fB0Prev := fB0; // 系数快照对齐首拍值，避免首拍误报变更沿 / align the snapshots to avoid a spurious change edge
    _fB1Prev := fB1; // 上拍 b1 快照对齐 / align the b1 snapshot
    _fB2Prev := fB2; // 上拍 b2 快照对齐 / align the b2 snapshot
    _fA1Prev := fA1; // 上拍 a1 快照对齐 / align the a1 snapshot
    _fA2Prev := fA2; // 上拍 a2 快照对齐 / align the a2 snapshot
END_IF
IF rtReset.Q THEN // 复位沿（作用域：清锁存 + 清滤波器状态，R311 声明）/ the reset edge with the declared scope
    _uLatch := 16#0000_0000; // 清故障码锁存（唯一的故障解除路径）/ clear the latched code, the only release path
    _fW1 := DL_BQ_ZERO; // 清状态 w1 / clear the state w1
    _fW2 := DL_BQ_ZERO; // 清状态 w2 / clear the state w2
END_IF
_bSatI := FALSE; // 钳位单拍内部位预清零 / preset the internal clamp bit false
_bCoefChg := FALSE; // 系数变更标记预清零 / preset the coefficient change flag false
_bCfgBadI := FALSE; // 组态非法标记预清零 / preset the configuration fault flag false

// 段 2｜八个浮点入参逐个点名有限闸（R272 全量枚举，含换算量与限值）/ segment 2, the full finiteness gate over all eight real pins
_bFinCoef := (fB0 = fB0) AND ((fB0 - fB0) = (fB0 - fB0))
          AND (fB1 = fB1) AND ((fB1 - fB1) = (fB1 - fB1))
          AND (fB2 = fB2) AND ((fB2 - fB2) = (fB2 - fB2))
          AND (fA1 = fA1) AND ((fA1 - fA1) = (fA1 - fA1))
          AND (fA2 = fA2) AND ((fA2 - fA2) = (fA2 - fA2)); // 五系数有限 / the five coefficients are finite
_bFinIn := (fIn = fIn) AND ((fIn - fIn) = (fIn - fIn)); // 输入有限 / the input is finite
_bFinDom := (fOutMin = fOutMin) AND ((fOutMin - fOutMin) = (fOutMin - fOutMin))
         AND (fOutMax = fOutMax) AND ((fOutMax - fOutMax) = (fOutMax - fOutMax)); // 限值有限 / the limits are finite

// 段 3｜稳定域闸与组态归因（边界一二，四个成因独立码，R190；v1.0.1 换 Jury 三条件）/ segment 3, the stability gate and the unique cause attribution
_bStable := (ABS(fA2) < DL_BQ_A2LIM) AND ((DL_BQ_ONE + fA1 + fA2) > DL_BQ_ZERO) AND ((DL_BQ_ONE - fA1 + fA2) > DL_BQ_ZERO); // Jury 三条件：|a2|<1 且 1+a1+a2>0 且 1−a1+a2>0 / the Jury three conditions, the magnitude of a2 below one and both half plane products positive
IF NOT _bFinCoef THEN // 成因一：系数非有限 / cause one, the coefficients are not finite
    _bCfgBadI := TRUE; // 置组态标记 / raise the configuration flag
    IF _uLatch = 16#0000_0000 THEN // 仅首因入锁存（后续成因不覆盖首因，R152）/ latch only the first cause so a later cause never overwrites it
        _uLatch := 16#0002_3736; // 故障级：系数非有限 / fault grade, the coefficients are not finite
    END_IF
ELSIF NOT _bFinDom THEN // 成因二：限值非有限 / cause two, the limits are not finite
    _bCfgBadI := TRUE; // 置组态标记 / raise the configuration flag
    IF _uLatch = 16#0000_0000 THEN // 仅首因入锁存 / latch only the first cause
        _uLatch := 16#0002_3737; // 故障级：输出钳位域非法 / fault grade, the clamp domain is illegal
    END_IF
ELSIF fOutMin > fOutMax THEN // 成因三：钳位域反序 / cause three, the clamp domain is reversed
    _bCfgBadI := TRUE; // 置组态标记 / raise the configuration flag
    IF _uLatch = 16#0000_0000 THEN // 仅首因入锁存 / latch only the first cause
        _uLatch := 16#0002_3737; // 故障级：输出钳位域非法（与限值非有限同一族，出口不可分）/ fault grade under the same clamp domain family
    END_IF
ELSIF NOT _bStable THEN // 成因四：越过 Jury 三条件稳定域（v1.0.1 换判据）/ cause four, the Jury conditions are exceeded
    _bCfgBadI := TRUE; // 置组态标记 / raise the configuration flag
    IF _uLatch = 16#0000_0000 THEN // 仅首因入锁存 / latch only the first cause
        _uLatch := 16#0002_3735; // 故障级：系数越过 Jury 三条件稳定域 / fault grade, the Jury conditions are exceeded
    END_IF
END_IF
IF (NOT _bFinIn) AND (_uLatch = 16#0000_0000) THEN // 成因五：输入非有限（不覆盖已有首因）/ cause five, the input is not finite, never overwriting an earlier cause
    _uLatch := 16#0002_373A; // 故障级：输入非有限 / fault grade, the input is not finite
END_IF

// 段 4｜使能失能分支最先消费：降级为安全值并清状态（边界五，FB33-4 声明行）/ segment 4, the disabled branch degrades to the safe value
IF NOT bEnable THEN // 失能 / disabled
    _fW1 := DL_BQ_ZERO; // 状态清零（失能即弃用历史）/ clear the state, the history is abandoned
    _fW2 := DL_BQ_ZERO; // 状态清零 / clear the state
    _fOutLast := DL_BQ_ZERO; // 输出归零（下游控制量失能须归零，非冻结末值）/ zero the output, a control quantity must fall to zero rather than freeze
    fOut := DL_BQ_ZERO; // 出口归零 [工程单位] / the outlet falls to zero
    bSat := FALSE; // 钳位位清零 / clear the clamp bit
    bCfgBad := (_uLatch <> 16#0000_0000); // 组态标记照实回放（与锁存同源）/ replay the configuration flag from the latch
    bValid := FALSE; // 输出不可用（安全值不是滤波结果，明示而非静默）/ mark the output unusable, a safe zero is not a filter result
    bError := (_uLatch <> 16#0000_0000); // 故障位照实回放 / replay the fault bit from the latch
    eErr := _uLatch; // 故障码锁存回放（信息级不参与失能分支）/ replay the latched code, informational codes do not apply while disabled
    RETURN; // 早退，不推进滤波 / early return without advancing the filter
END_IF

// 段 5｜组态故障或输入非有限：冻结最近有效输出，不推进状态（边界一二三，R273）/ segment 5, freeze on a fault without advancing the state
IF (_uLatch <> 16#0000_0000) OR _bCfgBadI OR (NOT _bFinIn) THEN // 任一故障相 / any fault phase
    IF (_fOutLast = _fOutLast) AND ((_fOutLast - _fOutLast) = (_fOutLast - _fOutLast)) THEN // 冻结源有限性闸（冻结只防推进不防污染，FB51-3）/ the frozen source finiteness gate
        fOut := _fOutLast; // 冻结最近有效输出 [工程单位] / freeze the last valid output
    ELSE // 冻结源自身被污染（理论上不可达）/ the frozen source itself is polluted, unreachable by theory
        _fOutLast := DL_BQ_ZERO; // 归零重建 / rebuild from zero
        fOut := DL_BQ_ZERO; // 出口归零 [工程单位] / the outlet falls to zero
    END_IF
    bSat := FALSE; // 钳位位清零 / clear the clamp bit
    bCfgBad := (_uLatch = 16#0002_3735) OR (_uLatch = 16#0002_3736) OR (_uLatch = 16#0002_3737); // bCfgBad 专指组态族三码，373A 输入坏不再复用（v1.0.1 修 R62-D5）/ the configuration flag now covers only the three configuration family codes, the input fault code no longer reuses it
    bValid := FALSE; // 输出不可用 / the output is not usable
    bError := TRUE; // 故障位置位 / raise the fault bit
    eErr := _uLatch; // 锁存码回放（不按当下输入重新推断，R152）/ replay the latched code instead of inferring from the current input
    RETURN; // 早退 / early return
END_IF

// 段 6｜系数变更沿：五系数任一 |新 − 旧| > 容差即清状态（边界三）/ segment 6, the coefficient change edge clears the state
IF (ABS(fB0 - _fB0Prev) > DL_BQ_EPS) OR (ABS(fB1 - _fB1Prev) > DL_BQ_EPS)
OR (ABS(fB2 - _fB2Prev) > DL_BQ_EPS) OR (ABS(fA1 - _fA1Prev) > DL_BQ_EPS)
OR (ABS(fA2 - _fA2Prev) > DL_BQ_EPS) THEN // 任一系数变更 / any coefficient changed
    _bCoefChg := TRUE; // 置变更标记（信息级 3739）/ raise the change flag for the informational code
    _fW1 := DL_BQ_ZERO; // 清状态 w1（防旧状态冲击新频响，保守处置）/ clear the state w1 to protect the new response from the old state
    _fW2 := DL_BQ_ZERO; // 清状态 w2 / clear the state w2
END_IF
_fB0Prev := fB0; // 系数快照推进 [−] / advance the b0 snapshot
_fB1Prev := fB1; // 系数快照推进 [−] / advance the b1 snapshot
_fB2Prev := fB2; // 系数快照推进 [−] / advance the b2 snapshot
_fA1Prev := fA1; // 系数快照推进 [−] / advance the a1 snapshot
_fA2Prev := fA2; // 系数快照推进 [−] / advance the a2 snapshot

// 段 7｜Direct Form I 差分方程（本拍中间量与输出）/ segment 7, the Direct Form I difference equation
_fW := fIn - (fA1 * _fW1) - (fA2 * _fW2); // 中间量 w = x − a1·w1 − a2·w2 [工程单位] / the intermediate w
_fY := (fB0 * _fW) + (fB1 * _fW1) + (fB2 * _fW2); // 输出 y = b0·w + b1·w1 + b2·w2 [工程单位] / the output y
_fW2 := _fW1; // 状态右移：w1 → w2 / shift the state, w1 becomes w2
_fW1 := _fW; // 状态推进：本拍 w → w1 / advance the state, the current w becomes w1

// 段 8｜输出钳位 + 抗 windup 状态回写（边界四）/ segment 8, the clamp with the anti windup state write back
IF _fY > fOutMax THEN // 超上界 / above the ceiling
    fOut := fOutMax; // 钳上界 [工程单位] / clamp to the ceiling
    _bSatI := TRUE; // 置钳位内部位 / raise the internal clamp bit
    _fW1 := fOutMax; // 状态回写（防积分式累积发散）[工程单位] / write the state back to stop the accumulating divergence
ELSIF _fY < fOutMin THEN // 超下界 / below the floor
    fOut := fOutMin; // 钳下界 [工程单位] / clamp to the floor
    _bSatI := TRUE; // 置钳位内部位 / raise the internal clamp bit
    _fW1 := fOutMin; // 状态回写 [工程单位] / write the state back
ELSE // 域内 / inside the domain
    fOut := _fY; // 直出输出 [工程单位] / pass the output through
END_IF

// 段 9｜全部内部量非有限复检：中间量或输出被污染即拒收并锁存（FB32-7 保持槽口径）/ segment 9, the finiteness recheck before the state is stored
IF (fOut <> fOut) OR ((fOut - fOut) <> (fOut - fOut))
OR (_fW <> _fW) OR ((_fW - _fW) <> (_fW - _fW)) THEN // 输出或中间量非有限（NaN 自反 / Inf 差值自减）/ a non finite output or intermediate, tested by reflexivity and by the self difference
    _fW1 := DL_BQ_ZERO; // 状态清零，禁污染物驻留 / clear the state so nothing polluted remains
    _fW2 := DL_BQ_ZERO; // 状态清零 / clear the state
    IF _uLatch = 16#0000_0000 THEN // 仅首因入锁存 / latch only the first cause
        _uLatch := 16#0002_373A; // 故障级：输入或中间量非有限 / fault grade, the input or the intermediate is not finite
    END_IF
    fOut := DL_BQ_ZERO; // 出口归零 [工程单位] / the outlet falls to zero
    bSat := FALSE; // 钳位位清零 / clear the clamp bit
    bCfgBad := FALSE; // 373A 属测量坏而非组态坏，bCfgBad 保持 FALSE（v1.0.1 修 R62-D5）/ the input fault is a measurement issue, the configuration flag stays false
    bValid := FALSE; // 输出不可用 / the output is not usable
    bError := TRUE; // 故障位置位 / raise the fault bit
    eErr := _uLatch; // 锁存码回放 / replay the latched code
    RETURN; // 早退 / early return
END_IF

// 段 10｜最近有效输出写回（写前已过非有限闸）/ segment 10, store the last valid output after the finiteness gate
_fOutLast := fOut; // 快照更新 [工程单位] / update the snapshot

// 段 11｜统一出口（单拍位映射 + 信息级重算，R187 / FB51-8）/ segment 11, the unified outlet
bSat := _bSatI; // 钳位位出口 / the clamp bit outlet
bCfgBad := (_uLatch <> 16#0000_0000); // 组态标记出口（与锁存同源，锁存型非单拍）/ the configuration flag outlet derived from the latch
bValid := TRUE; // 域内输出可用 / the in-domain output is usable
bError := (_uLatch <> 16#0000_0000); // 故障位出口（锁存派生，R99）/ the fault bit outlet derived from the latch
IF _uLatch <> 16#0000_0000 THEN // 故障锁存回放优先 / the latched fault replays first
    eErr := _uLatch; // 锁存码 [码] / the latched code
ELSIF _bSatI THEN // 输出钳位（信息级，逐拍重算）/ the output clamp, informational and recomputed each scan
    eErr := 16#0002_3738; // 信息级：本拍输出被钳位 / informational, the output was clamped on this scan
ELSIF _bCoefChg THEN // 系数变更（信息级，逐拍重算）/ the coefficient change, informational and recomputed each scan
    eErr := 16#0002_3739; // 信息级：系数变更沿触发状态清零 / informational, a coefficient change cleared the state
ELSE // 无事件 / no event
    eErr := 16#0000_0000; // 正常 / ok
END_IF
END_FUNCTION_BLOCK
